(* IEC 61131-3 sources: TetherPLC/tests/compat (part 4) *)

(* ---- tc3_eventlog_case.st ---- *)
// tc3_eventlog_case.st — e2e for tc3_eventlog (tplc-eventlog).
PROGRAM tc3_eventlog_case
VAR
    msg : FB_TcMessage;
    alm : FB_TcAlarm;
    qry : FB_TcEventQuery;
    lg : FB_TcEventLogger;
    eb : FB_TcEventBase;
    ar : FB_TcArguments;
    si : FB_TcSourceInfo;
    st : INT;
    mask AT %QD0 : UDINT;
    diag AT %QD4 : UDINT;
END_VAR
    diag := st;
    IF st = 0 THEN
        mask := 0;
        msg.nEventClass := 7; msg.nEventId := 42;
        msg.sText := 'pump on'; msg.nCmd := 1;  // send INFO
        st := 1;
    ELSIF st = 1 THEN
        IF msg.bDone AND msg.hEvent <> 0 THEN mask := mask OR 1; END_IF;
        msg.nCmd := 0;
        alm.nEventClass := 7; alm.nEventId := 99;
        alm.nSeverity := 3; alm.sText := 'temp high';
        st := 2;
    ELSIF st = 2 THEN
        alm.nCmd := 1;                          // raise alarm
        st := 3;
    ELSIF st = 3 THEN
        IF alm.bDone AND alm.bActive AND alm.nState = 1 THEN
            mask := mask OR 2;
        END_IF;
        alm.nCmd := 0;
        st := 4;
    ELSIF st = 4 THEN
        alm.nCmd := 2;                          // clear
        st := 5;
    ELSIF st = 5 THEN
        IF alm.bDone AND alm.nState = 2 AND alm.bActive THEN
            mask := mask OR 4;
        END_IF;
        alm.nCmd := 0;
        st := 6;
    ELSIF st = 6 THEN
        qry.nId := alm.hEvent; qry.nCmd := 4;  // query the entry
        st := 7;
    ELSIF st = 7 THEN
        IF qry.bDone AND qry.nState = 2 AND qry.nSeverity = 3
           AND qry.nEventId = 99 THEN
            mask := mask OR 8;
        END_IF;
        qry.nCmd := 0;
        st := 8;
    ELSIF st = 8 THEN
        alm.nCmd := 3;                          // confirm
        st := 9;
    ELSIF st = 9 THEN
        IF alm.bDone AND NOT alm.bActive THEN mask := mask OR 16; END_IF;
        alm.nCmd := 0;
        st := 10;
    ELSIF st = 10 THEN
        // wrong-state op must error: query the released id
        qry.nId := 255; qry.nCmd := 4;
        st := 11;
    ELSIF st = 11 THEN
        IF qry.bError THEN mask := mask OR 32; END_IF;
        qry.nCmd := 0;
        st := 12;
    ELSIF st = 12 THEN
        qry.nCmd := 5;                          // stats
        st := 13;
    ELSIF st = 13 THEN
        IF qry.bDone AND qry.nRaised = 2 AND qry.nCleared = 1
           AND qry.nConfirmed = 1 AND qry.nLive = 1 THEN
            mask := mask OR 64;
        END_IF;
        qry.nCmd := 0;
        st := 14;
    ELSIF st = 14 THEN
        // second alarm for the aggregate/logger surface
        alm.nEventClass := 8; alm.nEventId := 77;
        alm.nSeverity := 3; alm.sText := 'overtemp';
        alm.nCmd := 1;
        lg.nFilterClass := 8; lg.nFilterEid := 0;
        st := 15;
    ELSIF st = 15 THEN
        IF alm.bDone THEN mask := mask OR 128; END_IF;
        alm.nCmd := 0;
        lg.nCmd := 7;                           // IsAlarmRaised
        st := 16;
    ELSIF st = 16 THEN
        lg.nCmd := 0;
        IF lg.bFound AND lg.nEidOut = 77 AND lg.nState = 1 THEN
            mask := mask OR 256;
        END_IF;
        st := 17;
    ELSIF st = 17 THEN
        lg.nCmd := 8;                           // GetAlarm
        st := 18;
    ELSIF st = 18 THEN
        lg.nCmd := 0;
        IF lg.bFound AND FIND(lg.sTextOut, 'overtemp') > 0 THEN
            mask := mask OR 512;
        END_IF;
        // EqualsToEventEntry against journal id 2
        eb.EventClass := 8; eb.EventId := 77;
        eb.Severity := 3; eb.Text := 'overtemp';
        eb.cEntryId := 2; eb.nCmd := 3;
        st := 19;
    ELSIF st = 19 THEN
        eb.nCmd := 0;
        IF eb.bEqual THEN mask := mask OR 1024; END_IF;
        lg.nCmd := 9;                           // ExportLoggedEvents
        st := 20;
    ELSIF st = 20 THEN
        lg.nCmd := 0;
        IF LEN(lg.sExport) > 0
           AND FIND(lg.sExport, ';') > 0
           AND FIND(lg.sExport, 'overtemp') > 0 THEN
            mask := mask OR 2048;
        END_IF;
        st := 21;
    ELSIF st = 21 THEN
        lg.nCmd := 2;                           // ClearAlarms (class 8)
        st := 22;
    ELSIF st = 22 THEN
        lg.nCmd := 0;
        IF lg.nCount = 1 THEN mask := mask OR 4096; END_IF;
        st := 23;
    ELSIF st = 23 THEN
        lg.nCmd := 5;                           // ConfirmAlarms
        st := 24;
    ELSIF st = 24 THEN
        lg.nCmd := 0;
        IF lg.nCount = 1 THEN mask := mask OR 8192; END_IF;
        // third alarm for the *All* variants
        alm.nEventClass := 8; alm.nEventId := 78;
        alm.nSeverity := 3; alm.sText := 'vibration';
        alm.nCmd := 1;
        st := 25;
    ELSIF st = 25 THEN
        IF alm.bDone THEN mask := mask OR 16384; END_IF;
        alm.nCmd := 0;
        lg.nCmd := 3;                           // ClearAllAlarms
        st := 26;
    ELSIF st = 26 THEN
        lg.nCmd := 0;
        IF lg.nCount >= 1 THEN mask := mask OR 32768; END_IF;
        st := 27;
    ELSIF st = 27 THEN
        lg.nCmd := 6;                           // ConfirmAllAlarms
        st := 28;
    ELSIF st = 28 THEN
        lg.nCmd := 0;
        IF lg.nCount >= 1 THEN mask := mask OR 65536; END_IF;
        st := 29;
    ELSIF st = 29 THEN
        lg.nCmd := 4;                           // ClearLoggedEvents
        st := 30;
    ELSIF st = 30 THEN
        lg.nCmd := 0;
        IF lg.nCount >= 1 THEN mask := mask OR 131072; END_IF;
        // FB_TcEventBase comparisons + text requests
        eb.EventClass := 8; eb.EventId := 77;
        eb.Severity := 3; eb.Text := 'overtemp';
        eb.cClass := 8; eb.cId := 77; eb.cSev := 3;
        eb.cText := 'overtemp'; eb.nCmd := 1;   // EqualsTo
        st := 31;
    ELSIF st = 31 THEN
        eb.nCmd := 0;
        IF eb.bEqual THEN mask := mask OR 262144; END_IF;
        st := 32;
    ELSIF st = 32 THEN
        eb.nCmd := 2;                           // EqualsToEventClass
        st := 33;
    ELSIF st = 33 THEN
        eb.nCmd := 0;
        IF eb.bEqual THEN mask := mask OR 524288; END_IF;
        st := 34;
    ELSIF st = 34 THEN
        eb.nCmd := 5;                           // RequestEventClassName
        st := 35;
    ELSIF st = 35 THEN
        eb.nCmd := 0;
        IF FIND(eb.sOut, '8') = 1 THEN mask := mask OR 1048576; END_IF;
        st := 36;
    ELSIF st = 36 THEN
        eb.nCmd := 6;                           // RequestEventText
        st := 37;
    ELSIF st = 37 THEN
        eb.nCmd := 0;
        IF FIND(eb.sOut, 'overtemp') = 1 THEN
            mask := mask OR 2097152;
        END_IF;
        ar.nInt := 5; ar.nCmd := 1;             // AddInt
        st := 38;
    ELSIF st = 38 THEN
        ar.nCmd := 0;
        st := 39;
    ELSIF st = 39 THEN
        IF ar.nCount = 1 THEN mask := mask OR 4194304; END_IF;
        ar.sArg := 'hi'; ar.nCmd := 3;          // AddString
        st := 40;
    ELSIF st = 40 THEN
        ar.nCmd := 0;
        st := 41;
    ELSIF st = 41 THEN
        IF ar.nCount = 2 THEN mask := mask OR 8388608; END_IF;
        si.Name := 'main'; si.nCmd := 1;        // ExtendName
        st := 42;
    ELSIF st = 42 THEN
        si.nCmd := 0;
        IF si.Extended THEN mask := mask OR 16777216; END_IF;
        st := 43;
    ELSIF st = 43 THEN
        ar.nCmd := 5;                           // Clear args
        st := 44;
    ELSIF st = 44 THEN
        ar.nCmd := 0;
        st := 45;
    ELSIF st = 45 THEN
        IF ar.bEmpty THEN mask := mask OR 33554432; END_IF;
        st := 46;
    END_IF;
    msg(); alm(); qry(); lg(); eb(); ar(); si();
END_PROGRAM

(* ---- tc3_ftp_case.st ---- *)
PROGRAM Tc3FtpCase
VAR
    mask      AT %QD0   : DINT;
    st        : INT;
    conn      : FB_FTP_Connect;
    connBad   : FB_FTP_Connect;
    sz        : FB_FTP_Cmd;
    mkd       : FB_FTP_MkDir;
    dl        : FB_FTP_Download;
    ls        : FB_FTP_List;
    up        : FB_FTP_Upload;
    szUp      : FB_FTP_Cmd;
    fex       : FB_FTP_FileExists;
    dex       : FB_FTP_DirExists;
    rn        : FB_FTP_Rename;
    acc       : ARRAY[0..1023] OF BYTE;
    accLen    : UDINT;
    i         : UDINT;
    upData    : ARRAY[0..511] OF BYTE;
END_VAR

// autonomous FTP sequence against tests/compat/ftp_test_peer.py
// (TCP 2121, PASV). The peer serves /data.txt (68B), /bin.dat,
// dirs / and /pub. Each state's bExecute is high only while st
// equals its index, giving every FB one rising edge; bDone
// advances the machine.
upData[0] := 16#50; upData[1] := 16#4C; upData[2] := 16#43;   // 'P','L','C'
upData[3] := 16#20; upData[4] := 16#75; upData[5] := 16#70;   // ' ','u','p'
// "PLC upload payload 12345" = 24 bytes
upData[6] := 16#6C; upData[7] := 16#6F; upData[8] := 16#61;
upData[9] := 16#64; upData[10] := 16#20; upData[11] := 16#70;
upData[12] := 16#61; upData[13] := 16#79; upData[14] := 16#6C;
upData[15] := 16#6F; upData[16] := 16#61; upData[17] := 16#64;
upData[18] := 16#20; upData[19] := 16#31; upData[20] := 16#32;
upData[21] := 16#33; upData[22] := 16#34; upData[23] := 16#35;

conn(sHost := '127.0.0.1', nPort := 2121, sUser := 'u', sPass := 'p',
     bExecute := st = 0, bClose := st = 11, tTimeout := T#5S);
connBad(sHost := '127.0.0.1', nPort := 21999, sUser := 'u', sPass := 'p',
        bExecute := st = 10, bClose := FALSE, tTimeout := T#3S);
sz(nConnHandle := conn.nConnHandle, sCmd := 'SIZE /data.txt',
   bExecute := st = 1, tTimeout := T#3S);
mkd(nConnHandle := conn.nConnHandle, sPath := '/newdir',
    bExecute := st = 2, tTimeout := T#3S);
dl(nConnHandle := conn.nConnHandle, sRemotePath := '/data.txt',
   bExecute := st = 3, tTimeout := T#10S);
ls(nConnHandle := conn.nConnHandle, sRemotePath := '/',
   bExecute := st = 4, tTimeout := T#10S);
up(nConnHandle := conn.nConnHandle, sRemotePath := '/up.bin',
   nLen := 24, DATA := upData, bExecute := st = 5, tTimeout := T#10S);
szUp(nConnHandle := conn.nConnHandle, sCmd := 'SIZE /up.bin',
     bExecute := st = 6, tTimeout := T#3S);
fex(nConnHandle := conn.nConnHandle, sPath := '/data.txt',
    bExecute := st = 7, tTimeout := T#3S);
dex(nConnHandle := conn.nConnHandle, sPath := '/pub',
    bExecute := st = 8, tTimeout := T#10S);
rn(nConnHandle := conn.nConnHandle, sOldPath := '/data.txt',
   sNewPath := '/renamed.txt', bExecute := st = 9, tTimeout := T#10S);

// accumulate download chunks every scan while st = 3
IF dl.nChunk > 0 AND accLen + dl.nChunk <= 1024 THEN
    FOR i := 0 TO dl.nChunk - 1 DO
        acc[accLen + i] := dl.DATA[i];
    END_FOR;
    accLen := accLen + dl.nChunk;
END_IF;

IF st = 0 AND conn.bDone THEN
    // connect -> login completes, handle issued
    IF conn.nStatus = 1 AND conn.nConnHandle <> 0 AND
       conn.nErrId = 0 THEN
        mask := mask + 1;
    END_IF;
    st := 1;
ELSIF st = 1 AND sz.bDone THEN
    // SIZE /data.txt -> 213, text "68"
    IF sz.nStatus = 1 AND sz.nRespCode = 213 AND
       sz.sText = '68' THEN
        mask := mask + 2;
    END_IF;
    st := 2;
ELSIF st = 2 AND mkd.bDone THEN
    // MKD /newdir -> 257
    IF mkd.nStatus = 1 AND mkd.nRespCode = 257 THEN
        mask := mask + 4;
    END_IF;
    st := 3;
ELSIF st = 3 AND dl.bDone THEN
    // RETR /data.txt -> 68 bytes "Hello FTP World!\n"x4
    IF dl.nStatus = 1 AND dl.nTotal = 68 AND accLen = 68 AND
       acc[0] = 16#48 AND acc[16] = 16#0A THEN
        mask := mask + 8;
    END_IF;
    st := 4;
ELSIF st = 4 AND ls.bDone THEN
    // LIST / -> non-empty listing
    IF ls.nStatus = 1 AND ls.nTotal > 0 THEN
        mask := mask + 16;
    END_IF;
    st := 5;
ELSIF st = 5 AND up.bDone THEN
    // STOR /up.bin -> 226
    IF up.nStatus = 1 AND up.nRespCode = 226 THEN
        mask := mask + 32;
    END_IF;
    st := 6;
ELSIF st = 6 AND szUp.bDone THEN
    // SIZE /up.bin -> 213 "24"
    IF szUp.nStatus = 1 AND szUp.nRespCode = 213 AND
       szUp.sText = '24' THEN
        mask := mask + 64;
    END_IF;
    st := 7;
ELSIF st = 7 AND fex.bDone THEN
    // FileExists /data.txt -> SIZE 213
    IF fex.bExists AND fex.nRespCode = 213 THEN
        mask := mask + 128;
    END_IF;
    st := 8;
ELSIF st = 8 AND dex.bDone THEN
    // DirExists /pub -> LIST ok
    IF dex.bExists AND dex.nStatus = 1 THEN
        mask := mask + 256;
    END_IF;
    st := 9;
ELSIF st = 9 AND rn.bDone THEN
    // Rename /data.txt -> /renamed.txt: RNFR 350 + RNTO 250
    IF rn.nStatus = 1 AND rn.nRespCode = 250 AND NOT rn.bError THEN
        mask := mask + 512;
    END_IF;
    st := 10;
ELSIF st = 10 AND connBad.bDone THEN
    // refused connect -> STATUS 2
    IF connBad.nStatus = 2 THEN
        mask := mask + 1024;
    END_IF;
    st := 11;
ELSIF st = 11 AND conn.bDone THEN
    // CLOSE -> session torn down
    IF conn.nConnHandle = 0 THEN
        mask := mask + 2048;
    END_IF;
    st := 12;
END_IF;
END_PROGRAM

(* ---- tc3_iec870_case.st ---- *)
PROGRAM Tc3Iec870Case
VAR
    mask      AT %QD0   : DINT;
    st        : INT;
    i2        : INT;
    conn      : FB_IEC870_5_104Master;
    connBad   : FB_IEC870_5_104Master;
    snd       : FB_IEC870_SendAsdu;
    snd2      : FB_IEC870_SendAsdu;
    snd3      : FB_IEC870_SendAsdu;
    rcv       : FB_IEC870_RecvAsdu;
    pay1      : ARRAY[0..239] OF BYTE;
    pay2      : ARRAY[0..239] OF BYTE;
    pay3      : ARRAY[0..239] OF BYTE;
    gotSp     : BOOL;
    gotMe     : BOOL;
    gotCs     : BOOL;
    gotSc     : BOOL;
    // helper-test vars
    o64       : ARRAY[0..6] OF BYTE;
    tenc      : SYSTEMTIME_TO_CP56Time2a;
    tdec      : CP56Time2a_TO_SYSTEMTIME;
    hY        : UDINT;
    hMo       : UDINT;
    hD        : UDINT;
    hH        : UDINT;
    hMi       : UDINT;
    hS        : UDINT;
    hMs       : UDINT;
    hbIV      : BOOL;
    hbSU      : BOOL;
    hVer      : UDINT;
    hCot      : STRING[31];
    hTid      : STRING[31];
    hIoa      : UDINT;
    hSpi      : BOOL;
    hDpi      : UDINT;
    hVti      : UDINT;
END_VAR

// autonomous IEC 60870-5-104 exchange against
// tests/compat/iec870_test_peer.py (TCP 2480). The peer is a
// slave: STARTDT handshake, then answers C_IC_NA_1 with
// M_SP_NA_1 + M_ME_NA_1, echoes C_CS_NA_1, answers C_SC_NA_1
// with an act-con. rcv() runs every scan (consume-on-read);
// each send gets one EXEC edge via its own st step.
rcv(nConnHandle := conn.nConnHandle);
IF rcv.bDone THEN
    // M_SP_NA_1: type1 vsq1 cot3 ca1 payload = IOA(3)+SPI(1)
    IF rcv.nTypeId = 1 AND rcv.nLen = 4 AND
       rcv.pPayload[2] = 1 AND rcv.pPayload[3] = 1 THEN
        gotSp := TRUE;
    END_IF;
    // M_ME_NA_1: type9 payload = IOA(3)+int16+QDS = 6 bytes
    IF rcv.nTypeId = 9 AND rcv.nLen = 6 AND
       rcv.pPayload[2] = 2 AND rcv.pPayload[3] = 16#34 AND
       rcv.pPayload[4] = 16#12 AND rcv.pPayload[5] = 0 THEN
        gotMe := TRUE;
    END_IF;
    IF rcv.nTypeId = 103 THEN
        gotCs := TRUE;
    END_IF;
    IF rcv.nTypeId = 45 THEN
        gotSc := TRUE;
    END_IF;
END_IF;

conn(sHost := '127.0.0.1', nPort := 2480, nCA_Size := 2,
     nCOT_Size := 2, bExecute := st = 0, bClose := st = 10,
     tTimeout := T#3S);
connBad(sHost := '127.0.0.1', nPort := 19999,
        bExecute := st = 8, bClose := FALSE, tTimeout := T#3S);

// payload staging
// pay1: interrogation C_IC_NA_1 has no info objects (len 0)
// pay2: C_CS_NA_1 clock sync, CP56Time2a = 13:45:30.250
// octets0-1 = sec*1000+ms = 30250 -> LE16 0x762A = 42,118
pay2[0] := 42; pay2[1] := 118;
pay2[2] := 45;                  // minute=45
pay2[3] := 13;                  // hour=13
pay2[4] := 15;                  // day=15
pay2[5] := 6;                   // month=6
pay2[6] := 124;                 // year-1900 = 2024-1900 = 124
// pay3: C_SC_NA_1 single command IOA=5, SCS=on -> 4 bytes
pay3[0] := 0; pay3[1] := 0; pay3[2] := 5; pay3[3] := 16#80;

snd(nConnHandle := conn.nConnHandle, nTypeId := 100, nVSQ := 0,
    nCOT := 5, nCA := 1, nLen := 0, pPayload := pay1,
    bExecute := st = 1);
snd2(nConnHandle := conn.nConnHandle, nTypeId := 103, nVSQ := 0,
     nCOT := 6, nCA := 1, nLen := 7, pPayload := pay2,
     bExecute := st = 4);
snd3(nConnHandle := conn.nConnHandle, nTypeId := 45, nVSQ := 1,
     nCOT := 6, nCA := 1, nLen := 4, pPayload := pay3,
     bExecute := st = 6);

IF st = 0 AND conn.bDone THEN
    IF conn.nStatus = 1 AND conn.nConnHandle <> 0 AND
       conn.nSubState = 3 AND conn.nErrId = 0 THEN
        mask := mask + 1;
    END_IF;
    st := 1;
ELSIF st = 1 AND snd.bDone THEN
    IF snd.nStatus = 1 AND snd.nErrId = 0 THEN
        mask := mask + 2;
    END_IF;
    st := 2;
ELSIF st = 2 AND gotSp AND gotMe THEN
    mask := mask + 4;
    st := 3;
ELSIF st = 3 THEN
    st := 4;
ELSIF st = 4 AND snd2.bDone THEN
    IF snd2.nStatus = 1 AND snd2.nErrId = 0 THEN
        mask := mask + 8;
    END_IF;
    st := 5;
ELSIF st = 5 AND gotCs THEN
    mask := mask + 16;
    st := 6;
ELSIF st = 6 AND snd3.bDone THEN
    IF snd3.nStatus = 1 AND snd3.nErrId = 0 THEN
        mask := mask + 32;
    END_IF;
    st := 7;
ELSIF st = 7 AND gotSc THEN
    mask := mask + 64;
    st := 8;
ELSIF st = 8 AND connBad.bDone THEN
    IF connBad.nStatus = 2 THEN
        mask := mask + 128;
    END_IF;
    st := 9;
ELSIF st = 9 THEN
    // pure-helper checks (single scan)
    // CP56Time2a roundtrip: encode 2024-06-15 13:45:30.250.
    // FB VAR_OUTPUT stays on the instance; copy pTime -> o64.
    tenc(nYear := 2024, nMonth := 6, nDay := 15,
         nHour := 13, nMinute := 45, nSecond := 30, nMs := 250,
         bIV := FALSE, bSU := FALSE);
    i2 := 0;
    WHILE i2 < 7 DO
        o64[i2] := tenc.pTime[i2];
        i2 := i2 + 1;
    END_WHILE;
    tdec(pTime := o64);
    hY := tdec.nYear; hMo := tdec.nMonth; hD := tdec.nDay;
    hH := tdec.nHour; hMi := tdec.nMinute; hS := tdec.nSecond;
    hMs := tdec.nMs; hbIV := tdec.bIV; hbSU := tdec.bSU;
    IF hY = 2024 AND hMo = 6 AND hD = 15 AND hH = 13 AND
       hMi = 45 AND hS = 30 AND hMs = 250 AND NOT hbIV THEN
        mask := mask + 256;
    END_IF;
    hCot := ASDU101COT_TO_STRING(3);
    hTid := ASDU101TYPEID_TO_STRING(9);
    IF hCot = 'SPONTANEOUS' AND hTid = 'M_ME_NA_1' THEN
        mask := mask + 512;
    END_IF;
    hIoa := CP24IOA_TO_DWORD(0, 0, 5);
    hSpi := F_iecGetSPI(1);
    hDpi := F_iecGetDPI(2);
    hVti := F_iecIncVTI(32767);
    hVer := GetIec870_Version();
    IF hIoa = 5 AND hSpi AND hDpi = 2 AND hVti = 0 AND
       hVer = 16#0100 THEN
        mask := mask + 1024;
    END_IF;
    st := 10;
ELSIF st = 10 THEN
    // bClose := st = 10 gave one rising edge -> session closed
    IF conn.nConnHandle = 0 THEN
        mask := mask + 2048;
        st := 11;
    END_IF;
END_IF;

END_PROGRAM

(* ---- tc3_jsonxml_case.st ---- *)
// tc3_jsonxml_case.st — e2e for tc3_jsonxml (pure-ST JSON).
// Builds a flat JSON object with FB_JsonSaxWriter, checks the
// text shape with FIND (string equality is not usable here),
// then parses it back with FB_JsonSaxReader.
PROGRAM tc3_jsonxml_case
VAR
    w : FB_JsonSaxWriter;
    r : FB_JsonSaxReader;
    doc : STRING[255];
    st : INT;
    mask AT %QD0 : UDINT;
    diag AT %QD4 : UDINT;
END_VAR
    diag := st;
    IF st = 0 THEN
        mask := 0;
        w.nCmd := 1;                        // Begin
        st := 1;
    ELSIF st = 1 THEN
        w.nCmd := 0;
        w.sKey := 'sp'; w.fReal := 12.5;
        st := 2;
    ELSIF st = 2 THEN
        w.nCmd := 4;                        // AddReal sp
        st := 3;
    ELSIF st = 3 THEN
        w.nCmd := 0;
        w.sKey := 'n'; w.nInt := 7;
        st := 4;
    ELSIF st = 4 THEN
        w.nCmd := 3;                        // AddInt n
        st := 5;
    ELSIF st = 5 THEN
        w.nCmd := 0;
        w.sKey := 'ok'; w.bBool := TRUE;
        st := 6;
    ELSIF st = 6 THEN
        w.nCmd := 5;                        // AddBool ok
        st := 7;
    ELSIF st = 7 THEN
        w.nCmd := 0;
        w.sKey := 's'; w.sVal := 'abc';
        st := 8;
    ELSIF st = 8 THEN
        w.nCmd := 2;                        // AddString s
        st := 9;
    ELSIF st = 9 THEN
        w.nCmd := 0;
        w.sKey := 'z';
        st := 10;
    ELSIF st = 10 THEN
        w.nCmd := 6;                        // AddNull z
        st := 11;
    ELSIF st = 11 THEN
        w.nCmd := 0;                        // clear so End sees an edge
        st := 12;
    ELSIF st = 12 THEN
        w.nCmd := 7;                        // End
        st := 13;
    ELSIF st = 13 THEN
        w.nCmd := 0;
        doc := w.sDoc;
        // shape checks (FIND, not equality)
        IF FIND(doc, '{"sp":12.500') = 1 THEN mask := mask OR 1; END_IF;
        IF FIND(doc, ',"n":7') > 0 THEN mask := mask OR 2; END_IF;
        IF FIND(doc, ',"ok":true') > 0 THEN mask := mask OR 4; END_IF;
        IF FIND(doc, ',"s":"abc"') > 0 THEN mask := mask OR 8; END_IF;
        IF FIND(doc, ',"z":null}') > 0 THEN mask := mask OR 16; END_IF;
        r.sIn := doc;
        st := 14;
    ELSIF st = 14 THEN
        r.nCmd := 1;                        // Load
        st := 15;
    ELSIF st = 15 THEN
        r.nCmd := 0;
        r.sKey := 'n';
        st := 16;
    ELSIF st = 16 THEN
        r.nCmd := 3;                        // GetInt n
        st := 17;
    ELSIF st = 17 THEN
        r.nCmd := 0;
        IF r.bDone AND r.nOut = 7 THEN mask := mask OR 32; END_IF;
        r.sKey := 'sp';
        st := 18;
    ELSIF st = 18 THEN
        r.nCmd := 4;                        // GetReal sp
        st := 19;
    ELSIF st = 19 THEN
        r.nCmd := 0;
        IF r.bDone AND r.fOut = 12.5 THEN mask := mask OR 64; END_IF;
        r.sKey := 'ok';
        st := 20;
    ELSIF st = 20 THEN
        r.nCmd := 5;                        // GetBool ok
        st := 21;
    ELSIF st = 21 THEN
        r.nCmd := 0;
        IF r.bDone AND r.bOut THEN mask := mask OR 128; END_IF;
        r.sKey := 's';
        st := 22;
    ELSIF st = 22 THEN
        r.nCmd := 2;                        // GetString s
        st := 23;
    ELSIF st = 23 THEN
        r.nCmd := 0;
        IF r.bDone AND FIND(r.sOut, 'abc') = 1 THEN mask := mask OR 256; END_IF;
        r.sKey := 'missing';
        st := 24;
    ELSIF st = 24 THEN
        r.nCmd := 2;                        // absent key -> error
        st := 25;
    ELSIF st = 25 THEN
        r.nCmd := 0;
        IF r.bError THEN mask := mask OR 512; END_IF;
        w.nCmd := 1;                        // Begin nested doc
        st := 27;
    ELSIF st = 27 THEN
        w.nCmd := 0;
        w.sKey := 'dev';
        st := 28;
    ELSIF st = 28 THEN
        w.nCmd := 9;                        // ObjBegin dev
        st := 29;
    ELSIF st = 29 THEN
        w.nCmd := 0;
        w.sKey := 'name'; w.sVal := 'ax1';
        st := 30;
    ELSIF st = 30 THEN
        w.nCmd := 2;                        // AddString name
        st := 31;
    ELSIF st = 31 THEN
        w.nCmd := 0;
        w.sKey := 'spd'; w.nInt := 2;
        st := 32;
    ELSIF st = 32 THEN
        w.nCmd := 3;                        // AddInt spd
        st := 33;
    ELSIF st = 33 THEN
        w.nCmd := 0;
        st := 34;
    ELSIF st = 34 THEN
        w.nCmd := 11;                       // EndAny -> close dev
        st := 35;
    ELSIF st = 35 THEN
        w.nCmd := 0;
        w.sKey := 'axes';
        st := 36;
    ELSIF st = 36 THEN
        w.nCmd := 10;                       // ArrBegin axes
        st := 37;
    ELSIF st = 37 THEN
        w.nCmd := 0;
        w.sKey := ''; w.nInt := 0;
        st := 38;
    ELSIF st = 38 THEN
        w.nCmd := 3;                        // array elem 0 (scalar)
        st := 39;
    ELSIF st = 39 THEN
        w.nCmd := 0;
        w.sKey := '';
        st := 40;
    ELSIF st = 40 THEN
        w.nCmd := 9;                        // ObjBegin elem object
        st := 41;
    ELSIF st = 41 THEN
        w.nCmd := 0;
        w.sKey := 'id'; w.nInt := 0;
        st := 42;
    ELSIF st = 42 THEN
        w.nCmd := 3;                        // AddInt id
        st := 43;
    ELSIF st = 43 THEN
        w.nCmd := 0;
        w.sKey := 'pos'; w.nInt := 100;
        st := 44;
    ELSIF st = 44 THEN
        w.nCmd := 3;                        // AddInt pos
        st := 45;
    ELSIF st = 45 THEN
        w.nCmd := 0;
        st := 46;
    ELSIF st = 46 THEN
        w.nCmd := 11;                       // EndAny -> close elem obj
        st := 47;
    ELSIF st = 47 THEN
        w.nCmd := 0;
        w.sKey := '';
        st := 48;
    ELSIF st = 48 THEN
        w.nCmd := 9;                        // ObjBegin elem 1
        st := 49;
    ELSIF st = 49 THEN
        w.nCmd := 0;
        w.sKey := 'id'; w.nInt := 1;
        st := 50;
    ELSIF st = 50 THEN
        w.nCmd := 3;
        st := 51;
    ELSIF st = 51 THEN
        w.nCmd := 0;
        w.sKey := 'pos'; w.nInt := 250;
        st := 52;
    ELSIF st = 52 THEN
        w.nCmd := 3;
        st := 53;
    ELSIF st = 53 THEN
        w.nCmd := 0;
        st := 54;
    ELSIF st = 54 THEN
        w.nCmd := 11;                       // EndAny -> close elem 1
        st := 55;
    ELSIF st = 55 THEN
        w.nCmd := 0;
        st := 56;
    ELSIF st = 56 THEN
        w.nCmd := 11;                       // EndAny -> close axes
        st := 57;
    ELSIF st = 57 THEN
        w.nCmd := 0;
        st := 58;
    ELSIF st = 58 THEN
        w.nCmd := 7;                        // End root
        st := 59;
    ELSIF st = 59 THEN
        w.nCmd := 0;
        doc := w.sDoc;
        IF FIND(doc, '"dev":{"name":"ax1","spd":2}') > 0
        THEN mask := mask OR 1024; END_IF;
        IF FIND(doc, ',"axes":[0,{"id":0,"pos":100}') > 0
        THEN mask := mask OR 2048; END_IF;
        IF FIND(doc, '{"id":1,"pos":250}]}') > 0
        THEN mask := mask OR 4096; END_IF;
        r.sIn := doc;
        st := 60;
    ELSIF st = 60 THEN
        r.nCmd := 1;                        // Load
        st := 61;
    ELSIF st = 61 THEN
        r.nCmd := 0;
        r.sKey := 'dev.spd';
        st := 62;
    ELSIF st = 62 THEN
        r.nCmd := 3;                        // GetInt dev.spd
        st := 63;
    ELSIF st = 63 THEN
        r.nCmd := 0;
        IF r.bDone AND r.nOut = 2 THEN mask := mask OR 8192; END_IF;
        r.sKey := 'axes.2.pos';
        st := 64;
    ELSIF st = 64 THEN
        r.nCmd := 3;                        // GetInt axes.2.pos
        st := 65;
    ELSIF st = 65 THEN
        r.nCmd := 0;
        IF r.bDone AND r.nOut = 250 THEN mask := mask OR 16384; END_IF;
        r.sKey := 'dev';
        st := 66;
    ELSIF st = 66 THEN
        r.nCmd := 2;                        // GetString dev -> raw obj
        st := 67;
    ELSIF st = 67 THEN
        r.nCmd := 0;
        IF r.bDone AND FIND(r.sOut, '"name"') > 0
        THEN mask := mask OR 32768; END_IF;
        r.sKey := 'axes.0.id';
        st := 68;
    ELSIF st = 68 THEN
        r.nCmd := 3;                        // GetInt axes.0.id -> elem1 obj? no:
        st := 69;                           // axes.0 is scalar 0, .id fails
    ELSIF st = 69 THEN
        r.nCmd := 0;
        // axes.0 is the scalar element 0; path 'axes.0.id' must fail
        IF r.bError THEN mask := mask OR 65536; END_IF;
        st := 70;
    END_IF;
    w(); r();
END_PROGRAM

(* ---- tc3_jsonxml_dom_case.st ---- *)
// tc3_jsonxml_dom_case.st — e2e for FB_JsonDomParser: load a
// document, query the tree, serialize, build a tree, error path.
// Every command needs a dedicated arm state + a reap state that
// clears nCmd (edge detect prev=0).
PROGRAM tc3_jsonxml_dom_case
VAR
    d : FB_JsonDomParser;
    doc : STRING[255];
    hR : UDINT;
    hDev : UDINT;
    hId : UDINT;
    hAx : UDINT;
    hA1 : UDINT;
    hF : UDINT;
    hN : UDINT;
    hR2 : UDINT;
    st : INT;
    mask AT %QD0 : UDINT;
    diag AT %QD4 : UDINT;
END_VAR
    diag := st;
    IF st = 0 THEN
        mask := 0;
        doc := CONCAT('{"name":"ax1","dev":{"id":7,"spd":1.5}',
            ',"axes":[1,2,3],"flag":true,"note":null}');
        d.sIn := doc;
        d.nCmd := 1;                        // Load
        st := 1;
    ELSIF st = 1 THEN                        // reap Load
        d.nCmd := 0;
        IF d.bDone THEN mask := mask OR 1; END_IF;
        st := 2;
    ELSIF st = 2 THEN                        // arm Root
        d.nCmd := 3;
        st := 3;
    ELSIF st = 3 THEN                        // reap Root
        d.nCmd := 0;
        hR := d.hOut;
        IF hR <> 0 THEN mask := mask OR 2; END_IF;
        st := 4;
    ELSIF st = 4 THEN                        // arm NodeType root
        d.hNode := hR;
        d.nCmd := 7;
        st := 5;
    ELSIF st = 5 THEN                        // reap
        d.nCmd := 0;
        IF d.nOut = 1 THEN mask := mask OR 4; END_IF;
        st := 6;
    ELSIF st = 6 THEN                        // arm ChildCount root
        d.hNode := hR;
        d.nCmd := 6;
        st := 7;
    ELSIF st = 7 THEN                        // reap
        d.nCmd := 0;
        IF d.nOut = 5 THEN mask := mask OR 8; END_IF;
        st := 8;
    ELSIF st = 8 THEN                        // arm ChildByName dev
        d.hNode := hR; d.sKey := 'dev';
        d.nCmd := 5;
        st := 9;
    ELSIF st = 9 THEN                        // reap -> hDev
        d.nCmd := 0;
        hDev := d.hOut;
        IF hDev <> 0 THEN mask := mask OR 16; END_IF;
        st := 10;
    ELSIF st = 10 THEN                       // arm NodeType dev
        d.hNode := hDev;
        d.nCmd := 7;
        st := 11;
    ELSIF st = 11 THEN                       // reap
        d.nCmd := 0;
        IF d.nOut = 1 THEN mask := mask OR 32; END_IF;
        st := 12;
    ELSIF st = 12 THEN                       // arm ChildByName id
        d.hNode := hDev; d.sKey := 'id';
        d.nCmd := 5;
        st := 13;
    ELSIF st = 13 THEN                       // reap -> hId
        d.nCmd := 0;
        hId := d.hOut;
        st := 14;
    ELSIF st = 14 THEN                       // arm NodeText id
        d.hNode := hId;
        d.nCmd := 9;
        st := 15;
    ELSIF st = 15 THEN                       // reap
        d.nCmd := 0;
        IF FIND(d.sOut, '7') = 1 THEN
            mask := mask OR 64;
        END_IF;
        st := 16;
    ELSIF st = 16 THEN                       // arm ChildByName axes
        d.hNode := hR; d.sKey := 'axes';
        d.nCmd := 5;
        st := 17;
    ELSIF st = 17 THEN                       // reap -> hAx
        d.nCmd := 0;
        hAx := d.hOut;
        st := 18;
    ELSIF st = 18 THEN                       // arm ChildCount axes
        d.hNode := hAx;
        d.nCmd := 6;
        st := 19;
    ELSIF st = 19 THEN                       // reap
        d.nCmd := 0;
        IF d.nOut = 3 THEN mask := mask OR 128; END_IF;
        st := 20;
    ELSIF st = 20 THEN                       // arm Child axes[1]
        d.hNode := hAx; d.nIdx := 1;
        d.nCmd := 4;
        st := 21;
    ELSIF st = 21 THEN                       // reap -> hA1
        d.nCmd := 0;
        hA1 := d.hOut;
        st := 22;
    ELSIF st = 22 THEN                       // arm NodeText axes[1]
        d.hNode := hA1;
        d.nCmd := 9;
        st := 23;
    ELSIF st = 23 THEN                       // reap
        d.nCmd := 0;
        IF FIND(d.sOut, '2') = 1 THEN
            mask := mask OR 256;
        END_IF;
        st := 24;
    ELSIF st = 24 THEN                       // arm ChildByName flag
        d.hNode := hR; d.sKey := 'flag';
        d.nCmd := 5;
        st := 25;
    ELSIF st = 25 THEN                       // reap -> hF
        d.nCmd := 0;
        hF := d.hOut;
        st := 26;
    ELSIF st = 26 THEN                       // arm NodeText flag
        d.hNode := hF;
        d.nCmd := 9;
        st := 27;
    ELSIF st = 27 THEN                       // reap
        d.nCmd := 0;
        IF FIND(d.sOut, 'true') = 1 THEN
            mask := mask OR 512;
        END_IF;
        st := 28;
    ELSIF st = 28 THEN                       // arm ChildByName note
        d.hNode := hR; d.sKey := 'note';
        d.nCmd := 5;
        st := 29;
    ELSIF st = 29 THEN                       // reap -> hN
        d.nCmd := 0;
        hN := d.hOut;
        st := 30;
    ELSIF st = 30 THEN                       // arm NodeType note
        d.hNode := hN;
        d.nCmd := 7;
        st := 31;
    ELSIF st = 31 THEN                       // reap
        d.nCmd := 0;
        IF d.nOut = 6 THEN mask := mask OR 1024; END_IF;
        st := 32;
    ELSIF st = 32 THEN                       // arm NodeKey dev
        d.hNode := hDev;
        d.nCmd := 8;
        st := 33;
    ELSIF st = 33 THEN                       // reap
        d.nCmd := 0;
        IF FIND(d.sOut, 'dev') = 1 THEN
            mask := mask OR 2048;
        END_IF;
        st := 34;
    ELSIF st = 34 THEN                       // arm ToJson whole doc
        d.hNode := 0;
        d.nCmd := 10;
        st := 35;
    ELSIF st = 35 THEN                       // reap
        d.nCmd := 0;
        IF FIND(d.sOut, '"name":"ax1"') > 0
           AND FIND(d.sOut, '"axes":[1,2,3]') > 0 THEN
            mask := mask OR 4096;
        END_IF;
        st := 36;
    ELSIF st = 36 THEN                       // arm Clear
        d.nCmd := 2;
        st := 37;
    ELSIF st = 37 THEN                       // reap Clear
        d.nCmd := 0;
        st := 38;
    ELSIF st = 38 THEN                       // arm AppendObject r
        d.hNode := 0; d.sKey := 'r';
        d.nCmd := 11;
        st := 39;
    ELSIF st = 39 THEN                       // reap -> hR2
        d.nCmd := 0;
        hR2 := d.hOut;
        st := 40;
    ELSIF st = 40 THEN                       // arm AppendString a=v
        d.hNode := hR2; d.sKey := 'a'; d.sVal := 'v';
        d.nCmd := 13;
        st := 41;
    ELSIF st = 41 THEN                       // reap
        d.nCmd := 0;
        st := 42;
    ELSIF st = 42 THEN                       // arm AppendInt n=42
        d.hNode := hR2; d.sKey := 'n'; d.nInt := 42;
        d.nCmd := 14;
        st := 43;
    ELSIF st = 43 THEN                       // reap
        d.nCmd := 0;
        st := 44;
    ELSIF st = 44 THEN                       // arm ToJson built tree
        d.hNode := 0;
        d.nCmd := 10;
        st := 45;
    ELSIF st = 45 THEN                       // reap
        d.nCmd := 0;
        IF FIND(d.sOut, '{"a":"v","n":42}') = 1 THEN
            mask := mask OR 8192;
        END_IF;
        st := 46;
    ELSIF st = 46 THEN                       // arm malformed Load
        d.sIn := '{"a":}';
        d.nCmd := 1;
        st := 47;
    ELSIF st = 47 THEN                       // reap error
        d.nCmd := 0;
        IF d.bError THEN mask := mask OR 16384; END_IF;
        st := 48;
    END_IF;
    d();
END_PROGRAM

(* ---- tc3_jsonxml_pretty_case.st ---- *)
// tc3_jsonxml_pretty_case.st — e2e for FB_JsonSaxPrettyWriter:
// indented JSON output.  Every command needs a dedicated arm
// state and a reap state that clears nCmd (edge detect prev=0).
PROGRAM tc3_jsonxml_pretty_case
VAR
    pw : FB_JsonSaxPrettyWriter;
    st : INT;
    mask AT %QD0 : UDINT;
    diag AT %QD4 : UDINT;
END_VAR
    diag := st;
    IF st = 0 THEN
        mask := 0;
        pw.nInt := 2;
        pw.nCmd := 12;                       // SetIndent 2
        st := 1;
    ELSIF st = 1 THEN                        // reap
        pw.nCmd := 0;
        st := 2;
    ELSIF st = 2 THEN                        // arm Begin
        pw.nCmd := 1;
        st := 3;
    ELSIF st = 3 THEN                        // reap
        pw.nCmd := 0;
        st := 4;
    ELSIF st = 4 THEN                        // arm AddString name
        pw.sKey := 'name'; pw.sVal := 'ax1';
        pw.nCmd := 2;
        st := 5;
    ELSIF st = 5 THEN                        // reap
        pw.nCmd := 0;
        st := 6;
    ELSIF st = 6 THEN                        // arm ObjBegin dev
        pw.sKey := 'dev';
        pw.nCmd := 9;
        st := 7;
    ELSIF st = 7 THEN                        // reap
        pw.nCmd := 0;
        st := 8;
    ELSIF st = 8 THEN                        // arm AddInt id
        pw.sKey := 'id'; pw.nInt := 7;
        pw.nCmd := 3;
        st := 9;
    ELSIF st = 9 THEN                        // reap
        pw.nCmd := 0;
        st := 10;
    ELSIF st = 10 THEN                       // arm AddReal spd
        pw.sKey := 'spd'; pw.fReal := 1.5;
        pw.nCmd := 4;
        st := 11;
    ELSIF st = 11 THEN                       // reap
        pw.nCmd := 0;
        st := 12;
    ELSIF st = 12 THEN                       // arm AddBool en
        pw.sKey := 'en'; pw.bBool := TRUE;
        pw.nCmd := 5;
        st := 13;
    ELSIF st = 13 THEN                       // reap
        pw.nCmd := 0;
        st := 14;
    ELSIF st = 14 THEN                       // arm EndAny dev
        pw.nCmd := 11;
        st := 15;
    ELSIF st = 15 THEN                       // reap
        pw.nCmd := 0;
        st := 16;
    ELSIF st = 16 THEN                       // arm ArrBegin axes
        pw.sKey := 'axes';
        pw.nCmd := 10;
        st := 17;
    ELSIF st = 17 THEN                       // reap
        pw.nCmd := 0;
        st := 18;
    ELSIF st = 18 THEN                       // arm AddInt 1
        pw.nInt := 1;
        pw.nCmd := 3;
        st := 19;
    ELSIF st = 19 THEN                       // reap
        pw.nCmd := 0;
        st := 20;
    ELSIF st = 20 THEN                       // arm AddInt 2
        pw.nInt := 2;
        pw.nCmd := 3;
        st := 21;
    ELSIF st = 21 THEN                       // reap
        pw.nCmd := 0;
        st := 22;
    ELSIF st = 22 THEN                       // arm EndAny axes
        pw.nCmd := 11;
        st := 23;
    ELSIF st = 23 THEN                       // reap
        pw.nCmd := 0;
        st := 24;
    ELSIF st = 24 THEN                       // arm End root
        pw.nCmd := 7;
        st := 25;
    ELSIF st = 25 THEN                       // reap + checks
        pw.nCmd := 0;
        IF pw.bDone THEN mask := mask OR 1; END_IF;
        IF FIND(pw.sDoc, '"dev": {') > 0 THEN
            mask := mask OR 2;
        END_IF;
        IF FIND(pw.sDoc, '
    "id": 7') > 0 THEN
            mask := mask OR 4;
        END_IF;
        IF FIND(pw.sDoc, '"axes": [') > 0 THEN
            mask := mask OR 8;
        END_IF;
        IF FIND(pw.sDoc, '1.500') > 0 THEN
            mask := mask OR 16;
        END_IF;
        IF FIND(pw.sDoc, '
}') > 0 AND NOT pw.bError THEN
            mask := mask OR 32;
        END_IF;
        st := 26;
    END_IF;
    pw();
END_PROGRAM

(* ---- tc3_jsonxml_xml_case.st ---- *)
// tc3_jsonxml_xml_case.st — e2e for the XML half of tc3_jsonxml:
// FB_XmlDomParser load/query/serialize + build commands.
// Command FBs need a full scan with nCmd=0 between commands (edge
// detect on prev=0): every command gets a dedicated arm state, then
// a reap state that clears nCmd and reads the outputs.
PROGRAM tc3_jsonxml_xml_case
VAR
    x : FB_XmlDomParser;
    xdoc : STRING[1023];
    hRoot : UDINT;
    hDev : UDINT;
    hNm : UDINT;
    hPos : UDINT;
    hAx : UDINT;
    hTmp : UDINT;
    st : INT;
    mask AT %QD0 : UDINT;
    diag AT %QD4 : UDINT;
END_VAR
    diag := st;
    IF st = 0 THEN
        mask := 0;
        xdoc := CONCAT('<?xml version="1.0"?>',
            CONCAT('<root><dev id="ax1" unit="mm">',
            CONCAT('<name>motor</name><pos>100</pos></dev>',
            CONCAT('<axes><axis pos="1"/><axis pos="2"/>',
                   '<axis pos="3"/></axes></root>'))));
        x.sIn := xdoc; x.nCmd := 1;           // Load
        st := 1;
    // reap Load
    ELSIF st = 1 THEN
        x.nCmd := 0;
        IF x.bDone THEN mask := mask OR 1; END_IF;
        st := 2;
    // arm Root
    ELSIF st = 2 THEN
        x.nCmd := 3;
        st := 3;
    // reap Root
    ELSIF st = 3 THEN
        x.nCmd := 0;
        hRoot := x.hOut;
        IF hRoot <> 0 THEN mask := mask OR 2; END_IF;
        st := 4;
    // arm NodeName root
    ELSIF st = 4 THEN
        x.hNode := hRoot;
        x.nCmd := 6;
        st := 5;
    // reap NodeName
    ELSIF st = 5 THEN
        x.nCmd := 0;
        IF FIND(x.sOut, 'root') = 1 THEN
            mask := mask OR 4;
        END_IF;
        st := 6;
    // arm ChildByName dev
    ELSIF st = 6 THEN
        x.hNode := hRoot; x.sName := 'dev';
        x.nCmd := 5;
        st := 7;
    // reap -> hDev
    ELSIF st = 7 THEN
        x.nCmd := 0;
        hDev := x.hOut;
        IF hDev <> 0 THEN mask := mask OR 8; END_IF;
        st := 8;
    // arm AttrByName id
    ELSIF st = 8 THEN
        x.hNode := hDev; x.sName := 'id';
        x.nCmd := 10;
        st := 9;
    // reap attr id
    ELSIF st = 9 THEN
        x.nCmd := 0;
        IF FIND(x.sOut, 'ax1') = 1 THEN
            mask := mask OR 16;
        END_IF;
        st := 10;
    // arm AttrCount dev
    ELSIF st = 10 THEN
        x.hNode := hDev;
        x.nCmd := 8;
        st := 11;
    // reap AttrCount
    ELSIF st = 11 THEN
        x.nCmd := 0;
        IF x.nOut = 2 THEN mask := mask OR 32; END_IF;
        st := 12;
    // arm ChildByName name
    ELSIF st = 12 THEN
        x.hNode := hDev; x.sName := 'name';
        x.nCmd := 5;
        st := 13;
    // reap -> hNm
    ELSIF st = 13 THEN
        x.nCmd := 0;
        hNm := x.hOut;
        st := 14;
    // arm NodeText name
    ELSIF st = 14 THEN
        x.hNode := hNm;
        x.nCmd := 7;
        st := 15;
    // reap NodeText
    ELSIF st = 15 THEN
        x.nCmd := 0;
        IF FIND(x.sOut, 'motor') = 1 THEN
            mask := mask OR 64;
        END_IF;
        st := 16;
    // arm ChildByName pos
    ELSIF st = 16 THEN
        x.hNode := hDev; x.sName := 'pos';
        x.nCmd := 5;
        st := 17;
    // reap -> hPos
    ELSIF st = 17 THEN
        x.nCmd := 0;
        hPos := x.hOut;
        st := 18;
    // arm NodeText pos
    ELSIF st = 18 THEN
        x.hNode := hPos;
        x.nCmd := 7;
        st := 19;
    // reap NodeText pos
    ELSIF st = 19 THEN
        x.nCmd := 0;
        IF FIND(x.sOut, '100') = 1 THEN
            mask := mask OR 128;
        END_IF;
        st := 20;
    // arm ChildByName axes
    ELSIF st = 20 THEN
        x.hNode := hRoot; x.sName := 'axes';
        x.nCmd := 5;
        st := 21;
    // reap -> hAx
    ELSIF st = 21 THEN
        x.nCmd := 0;
        hAx := x.hOut;
        st := 22;
    // arm ChildCount axes
    ELSIF st = 22 THEN
        x.hNode := hAx;
        x.nCmd := 9;
        st := 23;
    // reap ChildCount
    ELSIF st = 23 THEN
        x.nCmd := 0;
        IF x.nOut = 3 THEN mask := mask OR 256; END_IF;
        st := 24;
    // arm Child axes[1] (0-based -> second axis)
    ELSIF st = 24 THEN
        x.hNode := hAx; x.nIdx := 1;
        x.nCmd := 4;
        st := 25;
    // reap -> hTmp
    ELSIF st = 25 THEN
        x.nCmd := 0;
        hTmp := x.hOut;
        st := 26;
    // arm AttrByName pos on axis2
    ELSIF st = 26 THEN
        x.hNode := hTmp; x.sName := 'pos';
        x.nCmd := 10;
        st := 27;
    // reap attr pos
    ELSIF st = 27 THEN
        x.nCmd := 0;
        IF FIND(x.sOut, '2') = 1 THEN
            mask := mask OR 512;
        END_IF;
        st := 28;
    // arm NodeXml dev
    ELSIF st = 28 THEN
        x.hNode := hDev;
        x.nCmd := 11;
        st := 29;
    // reap NodeXml
    ELSIF st = 29 THEN
        x.nCmd := 0;
        IF FIND(x.sOut, 'id="ax1"') > 0
           AND FIND(x.sOut, '<name>') > 0 THEN
            mask := mask OR 1024;
        END_IF;
        st := 30;
    // arm ToXml
    ELSIF st = 30 THEN
        x.hNode := 0;
        x.nCmd := 12;
        st := 31;
    // reap ToXml
    ELSIF st = 31 THEN
        x.nCmd := 0;
        IF FIND(x.sOut, '</root>') > 0
           AND FIND(x.sOut, '<axis') > 0 THEN
            mask := mask OR 2048;
        END_IF;
        st := 32;
    // arm Clear
    ELSIF st = 32 THEN
        x.nCmd := 2;
        st := 33;
    // reap Clear
    ELSIF st = 33 THEN
        x.nCmd := 0;
        st := 34;
    // arm AppendChild r under #doc
    ELSIF st = 34 THEN
        x.hNode := 0; x.sName := 'r';
        x.nCmd := 13;
        st := 35;
    // reap -> hRoot (new tree)
    ELSIF st = 35 THEN
        x.nCmd := 0;
        hRoot := x.hOut;
        st := 36;
    // arm AppendAttribute a=v on r
    ELSIF st = 36 THEN
        x.hNode := hRoot; x.sName := 'a'; x.sVal := 'v';
        x.nCmd := 14;
        st := 37;
    // reap attr
    ELSIF st = 37 THEN
        x.nCmd := 0;
        st := 38;
    // arm AppendChild c under r
    ELSIF st = 38 THEN
        x.hNode := hRoot; x.sName := 'c';
        x.nCmd := 13;
        st := 39;
    // reap -> hNm
    ELSIF st = 39 THEN
        x.nCmd := 0;
        hNm := x.hOut;
        st := 40;
    // arm AppendText hi on c
    ELSIF st = 40 THEN
        x.hNode := hNm; x.sVal := 'hi';
        x.nCmd := 15;
        st := 41;
    // reap text
    ELSIF st = 41 THEN
        x.nCmd := 0;
        st := 42;
    // arm ToXml of built tree
    ELSIF st = 42 THEN
        x.hNode := 0;
        x.nCmd := 12;
        st := 43;
    // reap ToXml
    ELSIF st = 43 THEN
        x.nCmd := 0;
        IF FIND(x.sOut, '<r a="v"><c>hi</c></r>') = 1 THEN
            mask := mask OR 4096;
        END_IF;
        st := 44;
    // arm malformed Load
    ELSIF st = 44 THEN
        x.sIn := '<a x></a>';
        x.nCmd := 1;
        st := 45;
    // reap error
    ELSIF st = 45 THEN
        x.nCmd := 0;
        IF x.bError THEN mask := mask OR 8192; END_IF;
        st := 46;
    END_IF;
    x();
END_PROGRAM

(* ---- tc3_mc2_ah_case.st ---- *)
// e2e for compat/tc3/tc3_mc2_ah.st — Tc3_MC2_AdvancedHoming:
// step search FBs (ref pulse, absolute switch, limit switch,
// block, block-lag), detection variants, finalizing FBs and a
// flying (passive) reference over a simulated axis.
// Mask bits (expected 0xFFFF):
//  0 axis created   1 powered        2 pos preset     3 refPulse
//  4 absSwitchDet   5 absSwitch      6 limitSwitch    7 block
//  8 blockDet       9 blockLag      10 homeDirect    11 finishHome
// 12 abortHome     13 flyingSwitch  14 errBadVel    15 errBadDir
PROGRAM Tc3Mc2AhCase
VAR
    mask   AT %QD0 : DINT;
    st     : INT;
    prevSt : INT;
    started: BOOL;
    pulse  : BOOL;

    ax     : FB_MotionAxis;
    rd     : FB_MotionAxis;
    axM    : UDINT;

    pwr    : MC_Power;
    sp     : MC_SetPosition;
    stp    : MC_Stop;
    mv     : MC_MoveVelocity;

    // homing FBs under test
    refPls : MC_StepReferencePulse;
    refPls2: MC_StepReferencePulse;
    refPls3: MC_StepReferencePulse;
    absDet : MC_StepAbsoluteSwitchDetection;
    absSw  : MC_StepAbsoluteSwitch;
    limSw  : MC_StepLimitSwitch;
    blk    : MC_StepBlock;
    blkDet : MC_StepBlockDetection;
    blkLag : MC_StepBlockLagBased;
    finH   : MC_FinishHoming;
    homeDir: MC_HomeDirect;
    abortH : MC_AbortHoming;
    flySw  : MC_StepReferenceFlyingSwitch;

    // shared MC_HomingParameter (flattened) state
    pStored : BOOL;
    pNcSMin : BOOL;  pNcSMax : BOOL;
    pNcSPosDiff : BOOL;  pNcSVeloDiff : BOOL;
    pNcAMin : BOOL;  pNcAMax : BOOL;
    pNcAPosDiff : BOOL;  pNcAVeloDiff : BOOL;
    pDrvSBip : LREAL;  pDrvSPos : LREAL;  pDrvSNeg : LREAL;
    pDrvABip : LREAL;  pDrvAPos : LREAL;  pDrvANeg : LREAL;

    // simulated reference signals (position-derived levels)
    dRef   : BOOL; dAbsD : BOOL; dAbsS : BOOL; dLim  : BOOL;
    dBlk   : BOOL; dBlkD : BOOL; dBlkL : BOOL; dHomeD : BOOL;
    dFin   : BOOL; dAbort: BOOL; dFly  : BOOL;
    sigZ   : BOOL;
    sigAbs : BOOL;
    sigLim : BOOL;
    sigFly : BOOL;

    posL   : LREAL;
    enSig  : BOOL;
    mvEx   : BOOL;
    spEx   : BOOL;
    stpEx  : BOOL;
    finEx  : BOOL;
    dirEx  : BOOL;
    abortEx: BOOL;
    flyEx  : BOOL;
    errEx  : BOOL;
    errEx2 : BOOL;
    refEx  : BOOL;
    absDetEx : BOOL;
    absSwEx  : BOOL;
    limSwEx  : BOOL;
    blkEx    : BOOL;
    blkDetEx : BOOL;
    blkLagEx : BOOL;
    homeDirEx: BOOL;
    errId1 : UDINT;
    errId2 : UDINT;
END_VAR

// ---- per-scan FB calls ----------------------------------------------
IF NOT started THEN
    pulse := TRUE; started := TRUE;
ELSIF st <> prevSt THEN
    pulse := TRUE;
ELSE
    pulse := FALSE;
END_IF;
prevSt := st;

IF axM <> 0 THEN
    rd.AXIS := axM; rd.OP := 6; rd();
END_IF;
posL := DINT_TO_LREAL(rd.POS_ACTUAL);

// reference signals derived from axis position
sigZ   := posL >= 5000.0;
sigAbs := posL >= 8000.0;
sigLim := posL <= -5000.0;
sigFly := posL >= 3000.0;

// execute pulses: launch stages, waits follow on the next stage
enSig := (st >= 1);
mvEx  := pulse AND (st = 38);
spEx  := pulse AND ((st = 2) OR (st = 6) OR (st = 10) OR (st = 14)
                    OR (st = 18) OR (st = 22) OR (st = 26));
stpEx := pulse AND (st = 42);
finEx := pulse AND (st = 33);
dirEx := pulse AND (st = 31);
abortEx := pulse AND (st = 35);
flyEx := pulse AND (st = 39);
errEx := pulse AND (st = 44);
errEx2 := pulse AND (st = 46);
refEx := pulse AND (st = 4);
absDetEx := pulse AND (st = 8);
absSwEx  := pulse AND (st = 12);
limSwEx  := pulse AND (st = 16);
blkEx    := pulse AND (st = 20);
blkDetEx := pulse AND (st = 24);
blkLagEx := pulse AND (st = 28);
homeDirEx:= dirEx;

pwr(Enable := enSig, Enable_Positive := TRUE, Enable_Negative := TRUE,
    Axis := axM);
sp(Execute := spEx, Position := 0, Mode := FALSE, Axis := axM);
stp(Execute := stpEx, Deceleration := 50000, Axis := axM);
mv(Execute := mvEx, ContinuousUpdate := FALSE, Velocity := 5000,
   Acceleration := 50000, Deceleration := 50000, Axis := axM);

// ---- homing FB calls (every scan; Execute is edge-driven inside) --
refPls(
       Execute := refEx,  Direction := 1,  SwitchMode := 3,
       RefLevel := sigZ,  Velocity := 20000.0,
       Acceleration := 50000.0,  Deceleration := 50000.0,  Jerk := 0.0,
       SetPosition := 100.0,  TimeLimit := T#0s,
       DistanceLimit := 50000.0,  TorqueLimit := 0.0,  BufferMode := 0,
       OptDisableDriveAccess := FALSE,
       OptEnableLagErrorDetection := FALSE,  Axis := axM,
       P_Stored := pStored,  P_NcSMin := pNcSMin,  P_NcSMax := pNcSMax,
       P_NcSPosDiff := pNcSPosDiff,  P_NcSVeloDiff := pNcSVeloDiff,
       P_NcAMin := pNcAMin,  P_NcAMax := pNcAMax,
       P_NcAPosDiff := pNcAPosDiff,  P_NcAVeloDiff := pNcAVeloDiff,
       P_DrvSBip := pDrvSBip,  P_DrvSPos := pDrvSPos,
       P_DrvSNeg := pDrvSNeg,  P_DrvABip := pDrvABip,
       P_DrvAPos := pDrvAPos,  P_DrvANeg := pDrvANeg);
absDet(
       Execute := absDetEx,  Direction := 3,  SwitchMode := 3,
       RefLevel := (posL <= -3000.0),  Velocity := 20000.0,
       Acceleration := 50000.0,  Deceleration := 50000.0,  Jerk := 0.0,
       TimeLimit := T#0s,  DistanceLimit := 50000.0,
       TorqueLimit := 0.0,  PositiveLimitSwitch := FALSE,
       NegativeLimitSwitch := FALSE,  BufferMode := 0,
       OptDisableDriveAccess := FALSE,
       OptEnableLagErrorDetection := FALSE,  Axis := axM,
       P_Stored := pStored,  P_NcSMin := pNcSMin,  P_NcSMax := pNcSMax,
       P_NcSPosDiff := pNcSPosDiff,  P_NcSVeloDiff := pNcSVeloDiff,
       P_NcAMin := pNcAMin,  P_NcAMax := pNcAMax,
       P_NcAPosDiff := pNcAPosDiff,  P_NcAVeloDiff := pNcAVeloDiff,
       P_DrvSBip := pDrvSBip,  P_DrvSPos := pDrvSPos,
       P_DrvSNeg := pDrvSNeg,  P_DrvABip := pDrvABip,
       P_DrvAPos := pDrvAPos,  P_DrvANeg := pDrvANeg);
absSw(
       Execute := absSwEx,  Direction := 1,  SwitchMode := 3,
       RefLevel := sigAbs,  Velocity := 20000.0,
       Acceleration := 50000.0,  Deceleration := 50000.0,  Jerk := 0.0,
       SetPosition := 500.0,  TimeLimit := T#0s,
       DistanceLimit := 50000.0,  TorqueLimit := 0.0,
       PositiveLimitSwitch := FALSE,  NegativeLimitSwitch := FALSE,
       BufferMode := 0,  OptDisableDriveAccess := FALSE,
       OptEnableLagErrorDetection := FALSE,  Axis := axM,
       P_Stored := pStored,  P_NcSMin := pNcSMin,  P_NcSMax := pNcSMax,
       P_NcSPosDiff := pNcSPosDiff,  P_NcSVeloDiff := pNcSVeloDiff,
       P_NcAMin := pNcAMin,  P_NcAMax := pNcAMax,
       P_NcAPosDiff := pNcAPosDiff,  P_NcAVeloDiff := pNcAVeloDiff,
       P_DrvSBip := pDrvSBip,  P_DrvSPos := pDrvSPos,
       P_DrvSNeg := pDrvSNeg,  P_DrvABip := pDrvABip,
       P_DrvAPos := pDrvAPos,  P_DrvANeg := pDrvANeg);
limSw(
       Execute := limSwEx,  Direction := 3,  LimitSwitchMode := 3,
       LimitSwitchLevel := sigLim,  Velocity := 20000.0,
       Acceleration := 50000.0,  Deceleration := 50000.0,  Jerk := 0.0,
       SetPosition := -500.0,  TimeLimit := T#0s,
       DistanceLimit := 50000.0,  TorqueLimit := 0.0,  BufferMode := 0,
       OptDisableDriveAccess := FALSE,
       OptEnableLagErrorDetection := FALSE,  Axis := axM,
       P_Stored := pStored,  P_NcSMin := pNcSMin,  P_NcSMax := pNcSMax,
       P_NcSPosDiff := pNcSPosDiff,  P_NcSVeloDiff := pNcSVeloDiff,
       P_NcAMin := pNcAMin,  P_NcAMax := pNcAMax,
       P_NcAPosDiff := pNcAPosDiff,  P_NcAVeloDiff := pNcAVeloDiff,
       P_DrvSBip := pDrvSBip,  P_DrvSPos := pDrvSPos,
       P_DrvSNeg := pDrvSNeg,  P_DrvABip := pDrvABip,
       P_DrvAPos := pDrvAPos,  P_DrvANeg := pDrvANeg);
blk(
       Execute := blkEx,  Direction := 1,  Velocity := 80000.0,
       Acceleration := 50000.0,  Deceleration := 50000.0,  Jerk := 0.0,
       SetPosition := 25000.0,  DetectionVelocityLimit := 800.0,
       DetectionVelocityTime := T#100ms,  TimeLimit := T#0s,
       DistanceLimit := 40000.0,  TorqueLimit := 0.0,
       TorqueTolerance := 0.0,  BufferMode := 0,
       OptDisableDriveAccess := FALSE,
       OptInstantLagReduction := FALSE,  Axis := axM,
       P_Stored := pStored,  P_NcSMin := pNcSMin,  P_NcSMax := pNcSMax,
       P_NcSPosDiff := pNcSPosDiff,  P_NcSVeloDiff := pNcSVeloDiff,
       P_NcAMin := pNcAMin,  P_NcAMax := pNcAMax,
       P_NcAPosDiff := pNcAPosDiff,  P_NcAVeloDiff := pNcAVeloDiff,
       P_DrvSBip := pDrvSBip,  P_DrvSPos := pDrvSPos,
       P_DrvSNeg := pDrvSNeg,  P_DrvABip := pDrvABip,
       P_DrvAPos := pDrvAPos,  P_DrvANeg := pDrvANeg);
blkDet(
       Execute := blkDetEx,  Direction := 3,  Velocity := 80000.0,
       Acceleration := 50000.0,  Deceleration := 50000.0,  Jerk := 0.0,
       DetectionVelocityLimit := 800.0,
       DetectionVelocityTime := T#100ms,  TimeLimit := T#0s,
       DistanceLimit := 40000.0,  TorqueLimit := 0.0,
       TorqueTolerance := 0.0,  BufferMode := 0,
       OptDisableDriveAccess := FALSE,
       OptInstantLagReduction := FALSE,  Axis := axM,
       P_Stored := pStored,  P_NcSMin := pNcSMin,  P_NcSMax := pNcSMax,
       P_NcSPosDiff := pNcSPosDiff,  P_NcSVeloDiff := pNcSVeloDiff,
       P_NcAMin := pNcAMin,  P_NcAMax := pNcAMax,
       P_NcAPosDiff := pNcAPosDiff,  P_NcAVeloDiff := pNcAVeloDiff,
       P_DrvSBip := pDrvSBip,  P_DrvSPos := pDrvSPos,
       P_DrvSNeg := pDrvSNeg,  P_DrvABip := pDrvABip,
       P_DrvAPos := pDrvAPos,  P_DrvANeg := pDrvANeg);
blkLag(
       Execute := blkLagEx,  Direction := 1,  Velocity := 80000.0,
       Acceleration := 50000.0,  Deceleration := 50000.0,  Jerk := 0.0,
       SetPosition := 20000.0,  DetectionVelocityLimit := 800.0,
       DetectionVelocityTime := T#100ms,  TimeLimit := T#0s,
       DistanceLimit := 40000.0,  TorqueLimit := 0.0,
       LagLimit := 1000.0,  BufferMode := 0,
       OptDisableDriveAccess := FALSE,
       OptInstantLagReduction := FALSE,  Axis := axM,
       P_Stored := pStored,  P_NcSMin := pNcSMin,  P_NcSMax := pNcSMax,
       P_NcSPosDiff := pNcSPosDiff,  P_NcSVeloDiff := pNcSVeloDiff,
       P_NcAMin := pNcAMin,  P_NcAMax := pNcAMax,
       P_NcAPosDiff := pNcAPosDiff,  P_NcAVeloDiff := pNcAVeloDiff,
       P_DrvSBip := pDrvSBip,  P_DrvSPos := pDrvSPos,
       P_DrvSNeg := pDrvSNeg,  P_DrvABip := pDrvABip,
       P_DrvAPos := pDrvAPos,  P_DrvANeg := pDrvANeg);
homeDir(
       Execute := homeDirEx,  SetPosition := 777.0,  BufferMode := 0,
       OptDisableDriveAccess := FALSE,  Axis := axM,
       P_Stored := pStored,  P_NcSMin := pNcSMin,  P_NcSMax := pNcSMax,
       P_NcSPosDiff := pNcSPosDiff,  P_NcSVeloDiff := pNcSVeloDiff,
       P_NcAMin := pNcAMin,  P_NcAMax := pNcAMax,
       P_NcAPosDiff := pNcAPosDiff,  P_NcAVeloDiff := pNcAVeloDiff,
       P_DrvSBip := pDrvSBip,  P_DrvSPos := pDrvSPos,
       P_DrvSNeg := pDrvSNeg,  P_DrvABip := pDrvABip,
       P_DrvAPos := pDrvAPos,  P_DrvANeg := pDrvANeg);
finH(
       Execute := finEx,  Distance := 500.0,  Velocity := 1000.0,
       Acceleration := 50000.0,  Deceleration := 50000.0,  Jerk := 0.0,
       BufferMode := 0,  OptDisableDriveAccess := FALSE,  Axis := axM,
       P_Stored := pStored,  P_NcSMin := pNcSMin,  P_NcSMax := pNcSMax,
       P_NcSPosDiff := pNcSPosDiff,  P_NcSVeloDiff := pNcSVeloDiff,
       P_NcAMin := pNcAMin,  P_NcAMax := pNcAMax,
       P_NcAPosDiff := pNcAPosDiff,  P_NcAVeloDiff := pNcAVeloDiff,
       P_DrvSBip := pDrvSBip,  P_DrvSPos := pDrvSPos,
       P_DrvSNeg := pDrvSNeg,  P_DrvABip := pDrvABip,
       P_DrvAPos := pDrvAPos,  P_DrvANeg := pDrvANeg);
abortH(
       Execute := abortEx,  OptDisableDriveAccess := FALSE,
       Axis := axM,  P_Stored := pStored,  P_NcSMin := pNcSMin,
       P_NcSMax := pNcSMax,  P_NcSPosDiff := pNcSPosDiff,
       P_NcSVeloDiff := pNcSVeloDiff,  P_NcAMin := pNcAMin,
       P_NcAMax := pNcAMax,  P_NcAPosDiff := pNcAPosDiff,
       P_NcAVeloDiff := pNcAVeloDiff,  P_DrvSBip := pDrvSBip,
       P_DrvSPos := pDrvSPos,  P_DrvSNeg := pDrvSNeg,
       P_DrvABip := pDrvABip,  P_DrvAPos := pDrvAPos,
       P_DrvANeg := pDrvANeg);
flySw(
       Execute := flyEx,  SwitchMode := 3,  RefLevel := sigFly,
       SetPosition := 4242.0,  TimeLimit := T#0s,
       DistanceLimit := 50000.0,  BufferMode := 0,  Axis := axM);
refPls2(
       Execute := errEx,  Direction := 1,  SwitchMode := 3,
       RefLevel := FALSE,  Velocity := 0.0,  Acceleration := 50000.0,
       Deceleration := 50000.0,  Jerk := 0.0,  SetPosition := 0.0,
       TimeLimit := T#0s,  DistanceLimit := 50000.0,
       TorqueLimit := 0.0,  BufferMode := 0,
       OptDisableDriveAccess := FALSE,
       OptEnableLagErrorDetection := FALSE,  Axis := axM,
       P_Stored := pStored,  P_NcSMin := pNcSMin,  P_NcSMax := pNcSMax,
       P_NcSPosDiff := pNcSPosDiff,  P_NcSVeloDiff := pNcSVeloDiff,
       P_NcAMin := pNcAMin,  P_NcAMax := pNcAMax,
       P_NcAPosDiff := pNcAPosDiff,  P_NcAVeloDiff := pNcAVeloDiff,
       P_DrvSBip := pDrvSBip,  P_DrvSPos := pDrvSPos,
       P_DrvSNeg := pDrvSNeg,  P_DrvABip := pDrvABip,
       P_DrvAPos := pDrvAPos,  P_DrvANeg := pDrvANeg);
refPls3(
       Execute := errEx2,  Direction := 9,  SwitchMode := 3,
       RefLevel := FALSE,  Velocity := 100.0,  Acceleration := 50000.0,
       Deceleration := 50000.0,  Jerk := 0.0,  SetPosition := 0.0,
       TimeLimit := T#0s,  DistanceLimit := 50000.0,
       TorqueLimit := 0.0,  BufferMode := 0,
       OptDisableDriveAccess := FALSE,
       OptEnableLagErrorDetection := FALSE,  Axis := axM,
       P_Stored := pStored,  P_NcSMin := pNcSMin,  P_NcSMax := pNcSMax,
       P_NcSPosDiff := pNcSPosDiff,  P_NcSVeloDiff := pNcSVeloDiff,
       P_NcAMin := pNcAMin,  P_NcAMax := pNcAMax,
       P_NcAPosDiff := pNcAPosDiff,  P_NcAVeloDiff := pNcAVeloDiff,
       P_DrvSBip := pDrvSBip,  P_DrvSPos := pDrvSPos,
       P_DrvSNeg := pDrvSNeg,  P_DrvABip := pDrvABip,
       P_DrvAPos := pDrvAPos,  P_DrvANeg := pDrvANeg);
// done latches (Done is a single-scan pulse)
IF refPls.Done THEN dRef := TRUE; END_IF;
IF absDet.Done THEN dAbsD := TRUE; END_IF;
IF absSw.Done THEN dAbsS := TRUE; END_IF;
IF limSw.Done THEN dLim := TRUE; END_IF;
IF blk.Done THEN dBlk := TRUE; END_IF;
IF blkDet.Done THEN dBlkD := TRUE; END_IF;
IF blkLag.Done THEN dBlkL := TRUE; END_IF;
IF homeDir.Done THEN dHomeD := TRUE; END_IF;
IF finH.Done THEN dFin := TRUE; END_IF;
IF abortH.Done THEN dAbort := TRUE; END_IF;
IF flySw.Done THEN dFly := TRUE; END_IF;

// latch single-scan error outputs
IF refPls2.Error THEN errId1 := refPls2.ErrorID; END_IF;
IF refPls3.Error THEN errId2 := refPls3.ErrorID; END_IF;

// ---- stages ----------------------------------------------------------
IF st = 0 THEN
    ax.UNITS_PER_REV := 1000;
    ax.MAX_VEL := 100000;
    ax.MAX_ACCEL := 200000;
    ax.MAX_DECEL := 200000;
    ax.POS_MIN := -20000;
    ax.POS_MAX := 30000;
    ax.HOME_OFFSET := 0;
    ax.FOLLOW_WINDOW := 3;
    ax.FLAGS := 1;
    ax.OP := 1; ax();
    IF ax.AXIS <> 0 THEN axM := ax.AXIS; END_IF;
    IF axM <> 0 THEN
        mask := mask + 1;                          // bit0
        // pos-limit objects (sim ext): needed on the IO backend
        // where axis create does not carry the config struct
        ax.AXIS := axM;
        ax.OP := 5; ax.INDEX := 16#200A; ax.VALUE := -20000; ax();
        ax.OP := 5; ax.INDEX := 16#200B; ax.VALUE := 30000;  ax();
        ax.OP := 5; ax.INDEX := 16#200C; ax.VALUE := 1;      ax();
    END_IF;
    st := 1;
ELSIF st = 1 THEN
    IF pwr.Status THEN mask := mask + 2; st := 2; END_IF;
ELSIF st = 2 THEN
    IF sp.Done THEN mask := mask + 4; st := 3; END_IF;
ELSIF st = 3 THEN st := 4;
ELSIF st = 4 THEN st := 5;
ELSIF st = 5 THEN
    IF dRef AND ABS(posL - 100.0) < 5.0 AND pStored = TRUE THEN
        mask := mask + 8; st := 6;
    END_IF;
ELSIF st = 6 THEN
    IF sp.Done THEN st := 7; END_IF;
ELSIF st = 7 THEN st := 8;
ELSIF st = 8 THEN st := 9;
ELSIF st = 9 THEN
    IF dAbsD AND absDet.RecordedPosition <= -2700.0
       AND absDet.RecordedPosition >= -3300.0 THEN
        mask := mask + 16; st := 10;
    END_IF;
ELSIF st = 10 THEN
    IF sp.Done THEN st := 11; END_IF;
ELSIF st = 11 THEN st := 12;
ELSIF st = 12 THEN st := 13;
ELSIF st = 13 THEN
    IF dAbsS AND ABS(posL - 500.0) < 5.0 THEN
        mask := mask + 32; st := 14;
    END_IF;
ELSIF st = 14 THEN
    IF sp.Done THEN st := 15; END_IF;
ELSIF st = 15 THEN st := 16;
ELSIF st = 16 THEN st := 17;
ELSIF st = 17 THEN
    IF dLim AND ABS(posL - (-500.0)) < 5.0 THEN
        mask := mask + 64; st := 18;
    END_IF;
ELSIF st = 18 THEN
    IF sp.Done THEN st := 19; END_IF;
ELSIF st = 19 THEN st := 20;
ELSIF st = 20 THEN st := 21;
ELSIF st = 21 THEN
    IF dBlk AND ABS(posL - 25000.0) < 5.0 THEN
        mask := mask + 128; st := 22;
    END_IF;
ELSIF st = 22 THEN
    IF sp.Done THEN st := 23; END_IF;
ELSIF st = 23 THEN st := 24;
ELSIF st = 24 THEN st := 25;
ELSIF st = 25 THEN
    IF dBlkD AND blkDet.RecordedPosition <= -19000.0
       AND blkDet.RecordedPosition >= -21000.0 THEN
        mask := mask + 256; st := 26;
    END_IF;
ELSIF st = 26 THEN
    IF sp.Done THEN st := 27; END_IF;
ELSIF st = 27 THEN st := 28;
ELSIF st = 28 THEN st := 29;
ELSIF st = 29 THEN
    IF dBlkL AND ABS(posL - 20000.0) < 5.0 THEN
        mask := mask + 512; st := 30;
    END_IF;
ELSIF st = 30 THEN st := 31;
ELSIF st = 31 THEN
    IF dHomeD AND ABS(posL - 777.0) < 5.0 THEN
        mask := mask + 1024; st := 32;
    END_IF;
ELSIF st = 32 THEN st := 33;
ELSIF st = 33 THEN
    IF dFin AND ABS(posL - 1277.0) < 60.0
       AND pStored = FALSE THEN
        mask := mask + 2048; st := 34;
    END_IF;
ELSIF st = 34 THEN st := 35;
ELSIF st = 35 THEN
    IF dAbort THEN mask := mask + 4096; st := 36; END_IF;
ELSIF st = 36 THEN st := 37;
ELSIF st = 37 THEN st := 38;
ELSIF st = 38 THEN st := 39;
ELSIF st = 39 THEN
    IF dFly AND posL >= 4242.0 AND posL <= 4800.0 THEN
        mask := mask + 8192; st := 40;
    END_IF;
ELSIF st = 40 THEN st := 41;
ELSIF st = 41 THEN st := 42;
ELSIF st = 42 THEN st := 43;
ELSIF st = 43 THEN st := 44;
ELSIF st = 44 THEN
    IF errId1 = 16#4B93 THEN mask := mask + 16384; END_IF;
    st := 45;
ELSIF st = 45 THEN st := 46;
ELSIF st = 46 THEN
    IF errId2 = 16#4B91 THEN mask := mask + 32768; END_IF;
    st := 47;
END_IF;
END_PROGRAM

(* ---- tc3_mc3cam_case.st ---- *)
PROGRAM Tc3Mc3CamCase
VAR
    mask   AT %QD0 : DINT;
    st     : INT;
    prevSt : INT;
    pulse  : BOOL;
    started : BOOL;
    axM    : UDINT;
    axS    : UDINT;
    crM    : FB_MotionAxis;
    crS    : FB_MotionAxis;
    rdM    : FB_MotionAxis;
    wrM    : FB_MotionAxis;
    wrS    : FB_MotionAxis;
    pwrM   : MC_Power;
    pwrS   : MC_Power;
    phA    : MC_PhasingAbsolute;
    phR    : MC_PhasingRelative;
    gip    : MC_GearInPos;
    hph    : MC_HaltPhasing;
    mpos   : DINT;
    spos   : DINT;
    dPhA   : BOOL;
    dPhR   : BOOL;
    dGip   : BOOL;
    dHph   : BOOL;
    gipOff : BOOL;
    phEx   : BOOL;
    relEx  : BOOL;
    gipEx  : BOOL;
    hphEx  : BOOL;
END_VAR

pulse := FALSE;
IF NOT started THEN
    pulse := TRUE; started := TRUE;
ELSIF st <> prevSt THEN
    pulse := TRUE;
END_IF;
prevSt := st;

// per-scan position reads (diagnostic only; FBs do their own)
IF axM <> 0 THEN
    rdM.AXIS := axM; rdM.OP := 4; rdM.INDEX := 16#6064; rdM();
    mpos := rdM.VALUE;
END_IF;
IF axS <> 0 THEN
    rdM.AXIS := axS; rdM.OP := 4; rdM.INDEX := 16#6064; rdM();
    spos := rdM.VALUE;
END_IF;

// Execute is edge-triggered inside each FB; level-held here
phEx  := st = 2;
relEx := st = 4;
gipEx := st = 5;
hphEx := st = 6;

phA(Execute := phEx, PhaseShift := 5000, Velocity := 50000,
    Acceleration := 0, Deceleration := 0, Jerk := 0,
    Master := axM, Slave := axS);
phR(Execute := relEx, PhaseShift := 2000, Velocity := 50000,
    Acceleration := 0, Deceleration := 0, Jerk := 0,
    Master := axM, Slave := axS);
gip(Execute := gipEx, RatioNumerator := 1, RatioDenominator := 1,
    Velocity := 50000, Acceleration := 0, Deceleration := 0,
    Jerk := 0, Master := axM, Slave := axS);
hph(Execute := hphEx, Deceleration := 0, Jerk := 0,
    Master := axM, Slave := axS);

IF phA.Done THEN dPhA := TRUE; END_IF;
IF phR.Done THEN dPhR := TRUE; END_IF;
IF gip.InSync THEN dGip := TRUE; END_IF;
IF hph.Done THEN dHph := TRUE; END_IF;

IF st = 0 THEN
    crM.UNITS_PER_REV := 1000; crM.MAX_VEL := 100000;
    crM.MAX_ACCEL := 200000; crM.MAX_DECEL := 200000;
    crM.POS_MIN := -100000; crM.POS_MAX := 100000;
    crM.HOME_OFFSET := 0; crM.FOLLOW_WINDOW := 3; crM.FLAGS := 1;
    crM.OP := 1; crM();
    IF crM.AXIS <> 0 THEN axM := crM.AXIS; END_IF;
    crS.UNITS_PER_REV := 1000; crS.MAX_VEL := 100000;
    crS.MAX_ACCEL := 200000; crS.MAX_DECEL := 200000;
    crS.POS_MIN := -100000; crS.POS_MAX := 100000;
    crS.HOME_OFFSET := 0; crS.FOLLOW_WINDOW := 3; crS.FLAGS := 1;
    crS.OP := 1; crS();
    IF crS.AXIS <> 0 THEN axS := crS.AXIS; END_IF;
    IF axM <> 0 AND axS <> 0 THEN mask := mask + 1; END_IF; // bit0
    st := 1;
ELSIF st = 1 THEN
    pwrM(Enable := TRUE, Enable_Positive := TRUE,
         Enable_Negative := TRUE, Axis := axM);
    pwrS(Enable := TRUE, Enable_Positive := TRUE,
         Enable_Negative := TRUE, Axis := axS);
    IF pwrM.Status AND pwrS.Status THEN
        mask := mask + 2; st := 2;                     // bit1
    END_IF;
ELSIF st = 2 THEN
    // master: PV mode, constant velocity 20000 u/s; phA edge fires
    wrM.AXIS := axM; wrM.OP := 5; wrM.INDEX := 16#6060;
    wrM.VALUE := 3; wrM();
    wrM.OP := 5; wrM.INDEX := 16#60FF; wrM.VALUE := 20000; wrM();
    st := 3;
ELSIF st = 3 THEN
    // absolute phasing: slave must reach masterPos + 5000
    IF dPhA THEN
        mask := mask + 4; st := 4;                     // bit2
    END_IF;
ELSIF st = 4 THEN
    // relative phasing: +2000 additional phase on top of offset0
    IF dPhR THEN
        mask := mask + 8; st := 5;                     // bit3
    END_IF;
ELSIF st = 5 THEN
    // offset the slave +2000 once; gear-in-position must pull it
    // back onto the anchored trajectory
    IF NOT gipOff THEN
        gipOff := TRUE;
        wrS.AXIS := axS; wrS.OP := 5; wrS.INDEX := 16#6064;
        wrS.VALUE := spos + 2000; wrS();
    END_IF;
    IF dGip THEN
        mask := mask + 16; st := 6;                    // bit4
    END_IF;
ELSIF st = 6 THEN
    // halt phasing: slave ramps to rest
    IF dHph THEN
        mask := mask + 32; st := 7;                    // bit5
    END_IF;
ELSIF st = 7 THEN
    // hold; expect written at final step
END_IF;
END_PROGRAM

(* ---- tc3_mc3camtbl_case.st ---- *)
// tc3_mc3camtbl_case.st — Tc3_Mc3Camming cam-table e2e over the
// tplc-cam service: FB_CamTable object creation + WritePt/Config
// edges, MC_CamTableSelect, MC_CamIn CSP coupling (slave tracks
// master+5000 through an identity cam table), MC_CamScaling offset
// update, MC_ReadCamInfo and MC_CamRemove. Mask 0xff (8 checks).
PROGRAM Tc3Mc3CamTblCase
VAR
    mask   AT %QD0 : DINT;
    st     : INT;
    prevSt : INT;
    pulse  : BOOL;
    started : BOOL;
    wrN    : INT;
    axM    : UDINT;
    axS    : UDINT;
    camH   : UDINT;
    crM    : FB_MotionAxis;
    crS    : FB_MotionAxis;
    wrM    : FB_MotionAxis;
    wrS    : FB_MotionAxis;
    pwrM   : MC_Power;
    pwrS   : MC_Power;
    tbl    : FB_CamTable;
    camI   : MC_CamIn;
    camS   : MC_CamScaling;
    camSel : MC_CamTableSelect;
    camR   : MC_CamRemove;
    camInfo: MC_ReadCamInfo;
    dSel   : BOOL;
    dScl   : BOOL;
    dRem   : BOOL;
    dInfo1 : BOOL;
    dInfo2 : BOOL;
    iFound : UDINT;
    iCam   : UDINT;
    iMaster: UDINT;
    jFound : UDINT;
    gapSeen : BOOL;
    selEx  : BOOL;
    camInEx: BOOL;
    camScEx: BOOL;
    camRemEx: BOOL;
    infoEx : BOOL;
END_VAR

pulse := FALSE;
IF NOT started THEN
    pulse := TRUE; started := TRUE;
ELSIF st <> prevSt THEN
    pulse := TRUE;
END_IF;
prevSt := st;

// ---- level inputs, computed before the FB calls ----
tbl.WritePt := FALSE; tbl.ClearTable := FALSE; tbl.Config := FALSE;
IF st = 3 THEN
    IF wrN = 0 THEN
        tbl.PtIndex := 0; tbl.PtMaster := 0.0; tbl.PtSlave := 0.0;
        tbl.WritePt := TRUE;
    ELSIF wrN = 2 THEN
        tbl.PtIndex := 1; tbl.PtMaster := 100000.0;
        tbl.PtSlave := 100000.0; tbl.WritePt := TRUE;
    ELSIF wrN = 3 THEN
        tbl.Config := TRUE; tbl.TableCount := 2;
        tbl.Periodic := FALSE; tbl.Continuity := 0;
    END_IF;
END_IF

selEx := st = 5;
camInEx := st = 6;
camScEx := st = 7;
camRemEx := st = 9;
infoEx := (st = 7) OR (st = 9);

camI(Execute := camInEx, Master := axM, Slave := axS,
     CamObject := camH, SlaveOffset := 5000.0);
camS(Execute := camScEx, Slave := axS, CamObject := camH,
     SlaveOffset := 8000.0);
camSel(Execute := selEx, CamRef := camH, Periodic := FALSE,
       ContinuityRequirement := 0, CamObjectIn := camH);
camR(Execute := camRemEx, Slave := axS, CamObject := camH);
camInfo(Execute := infoEx, Slave := axS);
tbl();

IF camSel.Done THEN dSel := TRUE; END_IF;
IF camS.Done THEN dScl := TRUE; END_IF;
IF camR.Done THEN dRem := TRUE; END_IF;
IF camInfo.Done THEN
    IF st = 7 THEN
        dInfo1 := TRUE;
        iFound := camInfo.NumberOfCouplingsFound;
        iCam := camInfo.CamHandle;
        iMaster := camInfo.MasterAxis;
    ELSIF st = 9 THEN
        dInfo2 := TRUE;
        jFound := camInfo.NumberOfCouplingsFound;
    END_IF;
END_IF;

IF st = 0 THEN
    crM.UNITS_PER_REV := 1000; crM.MAX_VEL := 100000;
    crM.MAX_ACCEL := 200000; crM.MAX_DECEL := 200000;
    crM.POS_MIN := -100000; crM.POS_MAX := 100000;
    crM.HOME_OFFSET := 0; crM.FOLLOW_WINDOW := 3; crM.FLAGS := 1;
    crM.OP := 1; crM();
    IF crM.AXIS <> 0 THEN axM := crM.AXIS; END_IF;
    crS.UNITS_PER_REV := 1000; crS.MAX_VEL := 100000;
    crS.MAX_ACCEL := 200000; crS.MAX_DECEL := 200000;
    crS.POS_MIN := -100000; crS.POS_MAX := 100000;
    crS.HOME_OFFSET := 0; crS.FOLLOW_WINDOW := 3; crS.FLAGS := 1;
    crS.OP := 1; crS();
    IF crS.AXIS <> 0 THEN axS := crS.AXIS; END_IF;
    IF axM <> 0 AND axS <> 0 THEN mask := mask + 1; END_IF; // bit0
    st := 1;
ELSIF st = 1 THEN
    pwrM(Enable := TRUE, Enable_Positive := TRUE,
         Enable_Negative := TRUE, Axis := axM);
    pwrS(Enable := TRUE, Enable_Positive := TRUE,
         Enable_Negative := TRUE, Axis := axS);
    IF pwrM.Status AND pwrS.Status THEN
        mask := mask + 2; st := 2;                     // bit1
    END_IF;
ELSIF st = 2 THEN
    // master PV move; slave into CSP mode for 0x607A streaming
    wrM.AXIS := axM; wrM.OP := 5; wrM.INDEX := 16#6060;
    wrM.VALUE := 3; wrM();
    wrM.OP := 5; wrM.INDEX := 16#60FF; wrM.VALUE := 5000; wrM();
    wrS.AXIS := axS; wrS.OP := 5; wrS.INDEX := 16#6060;
    wrS.VALUE := 8; wrS();
    wrN := 0;
    st := 3;
ELSIF st = 3 THEN
    // cam table point writes + config (wrN sequencer, ~5 scans)
    wrN := wrN + 1;
    IF wrN >= 5 THEN st := 4; END_IF;
ELSIF st = 4 THEN
    IF tbl.Handle <> 0 THEN
        camH := tbl.Handle;
        mask := mask + 4; st := 5;                     // bit2
    END_IF;
ELSIF st = 5 THEN
    IF dSel THEN
        mask := mask + 8; st := 6;                     // bit3
    END_IF;
ELSIF st = 6 THEN
    // MC_CamIn bound on entry; slave must converge to mpos+5000
    IF camI.InSync THEN
        mask := mask + 16; st := 7;                    // bit4
    END_IF;
ELSIF st = 7 THEN
    // scaling update + cam info read
    IF dScl AND dInfo1 THEN
        IF iFound = 1 AND iCam = camH AND iMaster = axM THEN
            mask := mask + 32;                        // bit5
        END_IF;
        st := 8;
    END_IF;
ELSIF st = 8 THEN
    // wait for the +3000 target jump to break sync, then re-converge
    IF NOT camI.InSync THEN gapSeen := TRUE; END_IF;
    IF gapSeen AND camI.InSync THEN
        mask := mask + 64; st := 9;                    // bit6
    END_IF;
ELSIF st = 9 THEN
    // cam remove + second info read must show no coupling
    IF dRem AND dInfo2 THEN
        IF jFound = 0 THEN
            mask := mask + 128;                       // bit7
        END_IF;
        st := 10;
    END_IF;
ELSIF st = 10 THEN
    // hold; expect written at final step
END_IF;
END_PROGRAM

(* ---- tc3_mc3ptp_case.st ---- *)
PROGRAM Tc3Mc3PtpCase
VAR
    mask   AT %QD0 : DINT;
    st     : INT;
    prevSt : INT;
    pulse  : BOOL;
    started : BOOL;
    axM    : UDINT;
    ax     : FB_MotionAxis;
    rd     : FB_MotionAxis;
    pwr    : MC_Power;
    rst    : MC_Reset;
    tq     : MC_ReadActualTorque;
    hwr    : MC_WriteHardwareParameter;
    hrr    : MC_ReadHardwareParameter;
    wfs    : MC_WaitForStableActualPosition;
    te     : MC_TriggerError;
    hs     : MC_SetHomingState;
    lc     : MC_LoadControl;
    esg    : MC_ActivateExternalSetpointGeneration;
    axErr  : MC_ReadAxisError;
    vel    : DINT;
END_VAR

// per-scan snapshot
IF axM <> 0 THEN
    rd.AXIS := axM; rd.OP := 6; rd();
    vel := rd.VEL_ACTUAL;
END_IF;

pulse := FALSE;
IF NOT started THEN
    pulse := TRUE; started := TRUE;
ELSIF st <> prevSt THEN
    pulse := TRUE;
END_IF;
prevSt := st;

IF st = 0 THEN
    ax.UNITS_PER_REV := 1000;
    ax.MAX_VEL := 100000;
    ax.MAX_ACCEL := 200000;
    ax.MAX_DECEL := 200000;
    ax.POS_MIN := -20000;
    ax.POS_MAX := 30000;
    ax.HOME_OFFSET := 0;
    ax.FOLLOW_WINDOW := 3;
    ax.FLAGS := 1;
    ax.OP := 1; ax();
    IF ax.AXIS <> 0 THEN axM := ax.AXIS; END_IF;
    IF axM <> 0 THEN mask := mask + 1; END_IF;   // bit0: create
    st := 1;
ELSIF st = 1 THEN
    pwr(Enable := TRUE, Enable_Positive := TRUE,
        Enable_Negative := TRUE, Axis := axM);
    IF pwr.Status THEN mask := mask + 2; st := 2; END_IF;  // bit1: power
ELSIF st = 2 THEN
    tq(Enable := TRUE, Axis := axM);
    hwr(Execute := pulse, ParameterNumber := 16#6065,
        Value := 5, Axis := axM);
    IF pulse AND hwr.Done AND tq.Valid THEN
        mask := mask + 4;                        // bit2: torque+hw wr
    END_IF;
    st := 3;
ELSIF st = 3 THEN
    hrr(Enable := TRUE, ParameterNumber := 16#6065, Axis := axM);
    IF hrr.Valid AND hrr.Value = 5 THEN
        mask := mask + 8;                        // bit3: hw param rd
    END_IF;
    st := 4;
ELSIF st = 4 THEN
    wfs(Execute := pulse, PositionWindow := 10,
        VelocityWindow := 1, Axis := axM);
    IF wfs.Done THEN mask := mask + 16; st := 5; END_IF;  // bit4: stable
ELSIF st = 5 THEN
    hs(Execute := pulse, HomingState := 1, Axis := axM);
    lc(Execute := pulse, Axis := axM);
    esg(Execute := pulse, Axis := axM);
    IF pulse AND hs.Done AND lc.Done AND esg.Done THEN
        mask := mask + 32;                       // bit5: no-op FBs
    END_IF;
    st := 6;
ELSIF st = 6 THEN
    te(Execute := pulse, ErrorCode := 4660, Axis := axM); // 0x1234
    IF pulse AND te.Done THEN mask := mask + 64; st := 7; END_IF; // bit6
ELSIF st = 7 THEN
    axErr(Enable := TRUE, Axis := axM);
    IF axErr.Valid AND axErr.AxisErrorID = 4660 THEN
        mask := mask + 128;                      // bit7: fault latched
    END_IF;
    rst(Execute := pulse, Axis := axM);
    IF pulse AND rst.Done THEN st := 8; END_IF;
ELSIF st = 8 THEN
    axErr(Enable := TRUE, Axis := axM);
    IF axErr.Valid AND axErr.AxisErrorID = 0 THEN
        mask := mask + 256;                      // bit8: fault cleared
    END_IF;
    st := 9;
ELSIF st = 9 THEN
    // hold; expect written at final step
END_IF;
END_PROGRAM

(* ---- tc3_mcgroup_case.st ---- *)
PROGRAM Tc3McGroupCase
VAR
    mask   AT %QD0 : DINT;
    st     : INT;
    prevSt : INT;
    cur    : INT;
    pulse  : BOOL;
    started : BOOL;
    grp    : UDINT;
    grpBad : UDINT;
    ax7    : UDINT;
    ax9    : UDINT;
    addA   : MC_AddAxisToGroup;
    addB   : MC_AddAxisToGroup;
    remA   : MC_RemoveAxisFromGroup;
    ungrp  : MC_UngroupAllAxes;
    enA    : MC_GroupEnable;
    enBad  : MC_GroupEnable;
    disA   : MC_GroupDisable;
    rstA   : MC_GroupReset;
    rs     : MC_GroupReadStatus;
    re     : MC_GroupReadError;
    so     : MC_GroupSetOverride;
    ss     : MC_GroupSetSetpointSource;
    ct     : MC_SetCoordinateTransform;
    ident  : UDINT;
    mg     : FB_McGroup;
    memOk  : BOOL;
END_VAR

cur := st;
pulse := (cur <> prevSt) OR NOT started;
started := TRUE;
prevSt := cur;

grp := 1;
grpBad := 2;
ax7 := 7;
ax9 := 9;
ident := UDINT_TO_IDENTINGROUP(0);
memOk := FALSE;

// Level-triggered readers: called every scan.
rs(Enable := TRUE, AxesGroup := grp);
re(Enable := TRUE, AxesGroup := grp);

// st0: add axis 7 to group 1 (ident 0)
IF cur = 0 THEN
    addA(Execute := pulse, IdentInGroup := ident,
         AxesGroup := grp, Axis := ax7);
    IF pulse AND addA.Done AND NOT addA.Error THEN
        mask := mask + 1;                       // bit0: add axis
    END_IF;
    st := 1;
// st1: status readback -> disabled, valid
ELSIF cur = 1 THEN
    IF rs.Valid AND rs.GroupDisabled THEN
        mask := mask + 2;                       // bit1: read status
    END_IF;
    st := 2;
// st2: enable group -> standby
ELSIF cur = 2 THEN
    enA(Execute := pulse, AxesGroup := grp);
    IF pulse AND enA.Done AND NOT enA.Error THEN
        mask := mask + 4;                       // bit2: enable done
    END_IF;
    st := 3;
// st3: status now standby + group error read valid
ELSIF cur = 3 THEN
    IF rs.GroupStandby AND re.Valid AND re.GroupErrorId = 0 THEN
        mask := mask + 8;                       // bit3: standby+err
    END_IF;
    st := 4;
// st4: enable empty group 2 -> error
ELSIF cur = 4 THEN
    enBad(Execute := pulse, AxesGroup := grpBad);
    IF pulse AND enBad.Error THEN
        mask := mask + 16;                      // bit4: empty enable err
    END_IF;
    st := 5;
// st5: override 150%
ELSIF cur = 5 THEN
    so(Execute := pulse, Enable := TRUE, VelFactor := 1.5,
       AxesGroup := grp);
    IF pulse AND so.Done AND
       ABS(so.OverrideActual - 1.5) < 0.001 THEN
        mask := mask + 32;                      // bit5: override
    END_IF;
    st := 6;
// st6: setpoint source MCS (2)
ELSIF cur = 6 THEN
    ss(Execute := pulse, SetpointSource := 2, AxesGroup := grp);
    IF pulse AND ss.Done AND NOT ss.Error THEN
        mask := mask + 64;                      // bit6: setpoint src
    END_IF;
    st := 7;
// st7: coordinate transform 3 -> active
ELSIF cur = 7 THEN
    ct(Execute := pulse, CoordTransform := 3, AxesGroup := grp);
    IF pulse AND ct.Done AND ct.Active AND NOT ct.Error THEN
        mask := mask + 128;                     // bit7: coord transform
    END_IF;
    st := 8;
// st8: membership readback via raw FB_McGroup OP10
ELSIF cur = 8 THEN
    mg.OP := 10; mg.GRP := grp; mg();
    IF mg.STATUS = 0 AND mg.NAXES = 1 AND mg.AXES[0] = 7 THEN
        memOk := TRUE;
        mask := mask + 256;                     // bit8: membership
    END_IF;
    st := 9;
// st9: disable group (membership changes need disabled state)
ELSIF cur = 9 THEN
    disA(Execute := pulse, AxesGroup := grp);
    IF pulse AND disA.Done THEN st := 10; END_IF;
// st10: add axis 9, remove axis 7 -> still 1 member (9)
ELSIF cur = 10 THEN
    addB(Execute := pulse, IdentInGroup := ident,
         AxesGroup := grp, Axis := ax9);
    remA(Execute := pulse, IdentInGroup := ident,
          AxesGroup := grp, Axis := ax7);
    IF pulse AND addB.Done AND remA.Done THEN st := 11; END_IF;
// st11: verify swap + ungroup all
ELSIF cur = 11 THEN
    mg.OP := 10; mg.GRP := grp; mg();
    IF mg.STATUS = 0 AND mg.NAXES = 1 AND mg.AXES[0] = 9 THEN
        mask := mask + 512;                     // bit9: swap member
    END_IF;
    ungrp(Execute := pulse, AxesGroup := grp);
    IF pulse AND ungrp.Done AND NOT ungrp.Error THEN
        mask := mask + 1024;                    // bit10: ungroup
    END_IF;
    st := 12;
// st12: group reset on fresh group
ELSIF cur = 12 THEN
    rstA(Execute := pulse, AxesGroup := grpBad);
    IF pulse AND rstA.Done THEN
        mask := mask + 2048;                    // bit11: reset
    END_IF;
    st := 13;
ELSIF cur = 13 THEN
    // hold; expect written at final step
END_IF;
END_PROGRAM

(* ---- tc3_mcgroup_stop_case.st ---- *)
// tc3_mcgroup_stop_case.st — Tc3_McCoordinatedMotion group motion
// e2e: two real axes grouped via MC_AddAxisToGroup, PV velocity
// moves, then MC_GroupStop (ramp to rest) and MC_GroupHalt
// (immediate disable) with per-axis VEL_ACTUAL verification.
// Mask 0x3f (6 checks).
PROGRAM Tc3McGroupStopCase
VAR
    mask   AT %QD0 : DINT;
    st     : INT;
    prevSt : INT;
    pulse  : BOOL;
    started : BOOL;
    dwell  : INT;
    grp    : UDINT := 1;
    axA    : UDINT;
    axB    : UDINT;
    crA    : FB_MotionAxis;
    crB    : FB_MotionAxis;
    rdA    : FB_MotionAxis;
    rdB    : FB_MotionAxis;
    wrA    : FB_MotionAxis;
    wrB    : FB_MotionAxis;
    pwrA   : MC_Power;
    pwrB   : MC_Power;
    addA   : MC_AddAxisToGroup;
    addB   : MC_AddAxisToGroup;
    gStop  : MC_GroupStop;
    gHalt  : MC_GroupHalt;
    vA     : DINT;
    vB     : DINT;
    dAddA  : BOOL;
    dAddB  : BOOL;
    dStop  : BOOL;
    dHalt  : BOOL;
    gStopEx: BOOL;
    gHaltEx: BOOL;
END_VAR

pulse := FALSE;
IF NOT started THEN
    pulse := TRUE; started := TRUE;
ELSIF st <> prevSt THEN
    pulse := TRUE; dwell := 0;
END_IF;
prevSt := st;

// per-scan velocity reads
IF axA <> 0 THEN
    rdA.AXIS := axA; rdA.OP := 3; rdA();
    rdA.OP := 4; rdA.INDEX := 16#606C; rdA(); vA := rdA.VALUE;
END_IF;
IF axB <> 0 THEN
    rdB.AXIS := axB; rdB.OP := 3; rdB();
    rdB.OP := 4; rdB.INDEX := 16#606C; rdB(); vB := rdB.VALUE;
END_IF;

gStopEx := st = 6;
gHaltEx := st = 10;
gStop(Execute := gStopEx, Deceleration := 1000.0, AxesGroup := grp);
gHalt(Execute := gHaltEx, AxesGroup := grp);

IF gStop.Done THEN dStop := TRUE; END_IF;
IF gHalt.Done THEN dHalt := TRUE; END_IF;

IF st = 0 THEN
    crA.UNITS_PER_REV := 1000; crA.MAX_VEL := 100000;
    crA.MAX_ACCEL := 200000; crA.MAX_DECEL := 200000;
    crA.POS_MIN := -100000; crA.POS_MAX := 100000;
    crA.HOME_OFFSET := 0; crA.FOLLOW_WINDOW := 3; crA.FLAGS := 1;
    crA.OP := 1; crA();
    IF crA.AXIS <> 0 THEN axA := crA.AXIS; END_IF;
    crB.UNITS_PER_REV := 1000; crB.MAX_VEL := 100000;
    crB.MAX_ACCEL := 200000; crB.MAX_DECEL := 200000;
    crB.POS_MIN := -100000; crB.POS_MAX := 100000;
    crB.HOME_OFFSET := 0; crB.FOLLOW_WINDOW := 3; crB.FLAGS := 1;
    crB.OP := 1; crB();
    IF crB.AXIS <> 0 THEN axB := crB.AXIS; END_IF;
    IF axA <> 0 AND axB <> 0 THEN mask := mask + 1; END_IF; // bit0
    st := 1;
ELSIF st = 1 THEN
    pwrA(Enable := TRUE, Enable_Positive := TRUE,
         Enable_Negative := TRUE, Axis := axA);
    pwrB(Enable := TRUE, Enable_Positive := TRUE,
         Enable_Negative := TRUE, Axis := axB);
    IF pwrA.Status AND pwrB.Status THEN
        mask := mask + 2; st := 2;                     // bit1
    END_IF;
ELSIF st = 2 THEN
    // add axis A to a fresh group (ensure creates the handle)
    addA(Execute := pulse, IdentInGroup := 0,
         AxesGroup := grp, Axis := axA);
    IF addA.Done THEN dAddA := TRUE; END_IF;
    IF dAddA THEN st := 3; END_IF;
ELSIF st = 3 THEN
    addB(Execute := pulse, IdentInGroup := 0,
         AxesGroup := grp, Axis := axB);
    IF addB.Done THEN dAddB := TRUE; END_IF;
    IF dAddB THEN
        mask := mask + 4; st := 4;                     // bit2
    END_IF;
ELSIF st = 4 THEN
    // both axes: PV mode, velocity 5000 u/s
    wrA.AXIS := axA; wrA.OP := 5; wrA.INDEX := 16#6060;
    wrA.VALUE := 3; wrA();
    wrA.OP := 5; wrA.INDEX := 16#60FF; wrA.VALUE := 5000; wrA();
    wrB.AXIS := axB; wrB.OP := 5; wrB.INDEX := 16#6060;
    wrB.VALUE := 3; wrB();
    wrB.OP := 5; wrB.INDEX := 16#60FF; wrB.VALUE := 5000; wrB();
    st := 5;
ELSIF st = 5 THEN
    // let both axes spin up, then confirm motion
    dwell := dwell + 1;
    IF dwell >= 15 THEN
        IF vA > 0 AND vB > 0 THEN
            mask := mask + 8;                         // bit3
        END_IF;
        st := 6;
    END_IF;
ELSIF st = 6 THEN
    // group stop: ramp to rest; Done implies all VEL_ACTUAL = 0
    IF dStop THEN
        mask := mask + 16; st := 7;                    // bit4
    END_IF;
ELSIF st = 7 THEN
    // restart both axes for the halt test
    wrA.AXIS := axA; wrA.OP := 5; wrA.INDEX := 16#6060;
    wrA.VALUE := 3; wrA();
    wrA.OP := 5; wrA.INDEX := 16#60FF; wrA.VALUE := 5000; wrA();
    wrB.AXIS := axB; wrB.OP := 5; wrB.INDEX := 16#6060;
    wrB.VALUE := 3; wrB();
    wrB.OP := 5; wrB.INDEX := 16#60FF; wrB.VALUE := 5000; wrB();
    st := 8;
ELSIF st = 8 THEN
    dwell := dwell + 1;
    IF dwell >= 15 THEN st := 10; END_IF;
ELSIF st = 10 THEN
    // group halt: immediate disable; Done implies all stopped
    IF dHalt THEN
        mask := mask + 32; st := 11;                   // bit5
    END_IF;
ELSIF st = 11 THEN
    // hold; expect written at final step
END_IF;
END_PROGRAM

(* ---- tc3_mcpath_case.st ---- *)
// tc3_mcpath_case.st — Tc3_McCoordinatedMotion path e2e: two real
// axes grouped, a 3-segment path (linear -> dwell -> linear)
// prepared through MC_MoveLinearAbsolutePreparation /
// MC_DwellTimePreparation, executed by MC_MovePath with per-scan
// 0x607A CSP streaming, final-position verification.
// Mask 0x3f (6 checks).
PROGRAM Tc3McPathCase
VAR
    mask   AT %QD0 : DINT;
    st     : INT;
    prevSt : INT;
    pulse  : BOOL;
    started : BOOL;
    grp    : UDINT := 1;
    pathH  : UDINT := 0;
    axA    : UDINT;
    axB    : UDINT;
    crA    : FB_MotionAxis;
    crB    : FB_MotionAxis;
    rdA    : FB_MotionAxis;
    rdB    : FB_MotionAxis;
    pwrA   : MC_Power;
    pwrB   : MC_Power;
    addA   : MC_AddAxisToGroup;
    addB   : MC_AddAxisToGroup;
    prep1  : MC_MoveLinearAbsolutePreparation;
    prepD  : MC_DwellTimePreparation;
    prepB  : MC_MoveBlendingPreparation;
    prepK  : MC_BlockerPreparation;
    relBlk : MC_ReleaseBlocker;
    blkSt  : MC_GroupReadBlockerStatus;
    trajRd : MC_GroupReadTrajectoryInformation;
    trafoPrep : MC_SetCoordinateTransformPreparation;
    setTrafo : MC_SetCoordinateTransform;
    mgRd   : FB_McGroup;
    prepC  : MC_MoveCircularAbsolutePreparation;
    prep2  : MC_MoveDirectPreparation;
    mvPath : MC_MovePath;
    pos1   : ARRAY[0..15] OF LREAL;
    pos2   : ARRAY[0..15] OF LREAL;
    auxC   : ARRAY[0..15] OF LREAL;
    endC   : ARRAY[0..15] OF LREAL;
    transP : ARRAY[0..15] OF LREAL;
    dAddA  : BOOL;
    dAddB  : BOOL;
    dPrep1 : BOOL;
    dPrepD : BOOL;
    dPrep2 : BOOL;
    dPath  : BOOL;
    busySeen : BOOL;
    gotBusy : BOOL;
    gotPos  : BOOL;
    sawBlocked : BOOL;
    sawTraj : BOOL;
    coordNow : UDINT;
    mCnt   : INT;
    dRel   : BOOL;
    pA     : DINT;
    pB     : DINT;
END_VAR

pulse := FALSE;
IF NOT started THEN
    pulse := TRUE; started := TRUE;
ELSIF st <> prevSt THEN
    pulse := TRUE;
END_IF;
prevSt := st;

// per-scan position reads
IF axA <> 0 THEN
    rdA.AXIS := axA; rdA.OP := 4; rdA.INDEX := 16#6064; rdA(); pA := rdA.VALUE;
END_IF;
IF axB <> 0 THEN
    rdB.AXIS := axB; rdB.OP := 4; rdB.INDEX := 16#6064; rdB(); pB := rdB.VALUE;
END_IF;

mvPath(Execute := st = 8, AxesGroup := grp, PathData := pathH);
IF mvPath.Busy THEN busySeen := TRUE; END_IF;
IF mvPath.Done THEN dPath := TRUE; END_IF;

IF st = 0 THEN
    crA.UNITS_PER_REV := 1000; crA.MAX_VEL := 100000;
    crA.MAX_ACCEL := 200000; crA.MAX_DECEL := 200000;
    crA.POS_MIN := -100000; crA.POS_MAX := 100000;
    crA.HOME_OFFSET := 0; crA.FOLLOW_WINDOW := 3; crA.FLAGS := 1;
    crA.OP := 1; crA();
    IF crA.AXIS <> 0 THEN axA := crA.AXIS; END_IF;
    crB.UNITS_PER_REV := 1000; crB.MAX_VEL := 100000;
    crB.MAX_ACCEL := 200000; crB.MAX_DECEL := 200000;
    crB.POS_MIN := -100000; crB.POS_MAX := 100000;
    crB.HOME_OFFSET := 0; crB.FOLLOW_WINDOW := 3; crB.FLAGS := 1;
    crB.OP := 1; crB();
    IF crB.AXIS <> 0 THEN axB := crB.AXIS; END_IF;
    IF axA <> 0 AND axB <> 0 THEN mask := mask + 1; END_IF; // bit0
    st := 1;
ELSIF st = 1 THEN
    pwrA(Enable := TRUE, Enable_Positive := TRUE,
         Enable_Negative := TRUE, Axis := axA);
    pwrB(Enable := TRUE, Enable_Positive := TRUE,
         Enable_Negative := TRUE, Axis := axB);
    IF pwrA.Status AND pwrB.Status THEN
        mask := mask + 2; st := 2;                     // bit1
    END_IF;
ELSIF st = 2 THEN
    addA(Execute := pulse, IdentInGroup := 0,
         AxesGroup := grp, Axis := axA);
    IF addA.Done THEN dAddA := TRUE; END_IF;
    IF dAddA THEN st := 3; END_IF;
ELSIF st = 3 THEN
    addB(Execute := pulse, IdentInGroup := 0,
         AxesGroup := grp, Axis := axB);
    setTrafo(Execute := pulse, CoordTransform := 3,
             AxesGroup := grp);
    IF addB.Done THEN dAddB := TRUE; END_IF;
    IF dAddB THEN
        mask := mask + 4; st := 4;                     // bit2
    END_IF;
ELSIF st = 4 THEN
    // segment 1: linear to (1000, 0)
    pos1[0] := 1000.0; pos1[1] := 0.0;
    prep1(Execute := pulse, Position := pos1, PositionCount := 2,
          Velocity := 20000.0, Acceleration := 50000.0,
          Deceleration := 50000.0, Jerk := 0.0, BufferMode := 1,
          PathData := pathH);
    IF prep1.Error THEN mask := mask + 256; END_IF;
    IF NOT prep1.Error THEN dPrep1 := TRUE; END_IF;
    IF dPrep1 THEN st := 5; END_IF;
ELSIF st = 5 THEN
    // segment 2: circular, center (0,0), end (0,1000), CCW
    auxC[0] := 0.0; auxC[1] := 0.0;
    endC[0] := 0.0; endC[1] := 1000.0;
    prepC(Execute := pulse, CircMode := 1,
          AuxPoint := auxC, AuxPointCount := 2,
          EndPoint := endC, EndPointCount := 2,
          PathChoice := 1, Velocity := 20000.0,
          Acceleration := 50000.0, Deceleration := 50000.0,
          Jerk := 0.0, BufferMode := 1, PathData := pathH);
    IF prepC.Error THEN mask := mask + 256; END_IF;
    IF NOT prepC.Error THEN dPrepD := TRUE; END_IF;
    IF dPrepD THEN st := 6; END_IF;
ELSIF st = 6 THEN
    // segment 3: dwell 200 ms, then a 150 ms blend junction
    prepD(Execute := pulse, DwellTime := 200, BufferMode := 1,
          PathData := pathH);
    transP[0] := 150.0;
    prepB(Execute := pulse, Velocity := 20000.0,
          Acceleration := 50000.0, Deceleration := 50000.0,
          Jerk := 0.0, BufferMode := 1, TransitionMode := 0,
          TransitionParameter := transP,
          TransitionParameterCount := 1, InvokeId := 0,
          PathData := pathH);
    IF prepD.Error OR prepB.Error THEN mask := mask + 256; END_IF;
    IF NOT prepD.Error AND NOT prepB.Error THEN st := 7; END_IF;
ELSIF st = 7 THEN
    // transform marker -> coord 9, blocker gate id 7, linear
    trafoPrep(PathData := pathH, CoordTransform := 9);
    prepK(Execute := pulse, BlockerId := 7, BufferMode := 1,
          PathData := pathH);
    pos2[0] := 2000.0; pos2[1] := 2000.0;
    prep2(Execute := pulse, Position := pos2, PositionCount := 2,
          Velocity := 20000.0, Acceleration := 50000.0,
          Deceleration := 50000.0, Jerk := 0.0, BufferMode := 1,
          PathData := pathH);
    IF prepK.Error OR prep2.Error THEN mask := mask + 256; END_IF;
    IF NOT prepK.Error AND NOT prep2.Error THEN dPrep2 := TRUE; END_IF;
    IF dPrep2 THEN
        // 6 segments prepared on a live path handle
        IF pathH <> 0 THEN mask := mask + 8; END_IF;   // bit3
        st := 8;
    END_IF;
ELSIF st = 8 THEN
    // path running; blocker status polled, release after ~1.2 s
    blkSt(Enable := TRUE, AxesGroup := grp);
    IF blkSt.Blocked THEN sawBlocked := TRUE; END_IF;
    trajRd(Enable := TRUE, AxesGroup := grp);
    IF trajRd.Valid AND trajRd.EntryCount >= 3 THEN
        sawTraj := TRUE;
    END_IF;
    IF busySeen THEN gotBusy := TRUE; END_IF;
    mCnt := mCnt + 1;
    IF mCnt >= 120 THEN st := 9; END_IF;
ELSIF st = 9 THEN
    // release the blocker gate
    relBlk(Execute := pulse, BlockerId := 7, AxesGroup := grp);
    IF relBlk.Done THEN dRel := TRUE; END_IF;
    IF dRel THEN st := 10; END_IF;
ELSIF st = 10 THEN
    // path resumes and finishes
    IF dPath THEN
        // final positions near (2000, 2000), tolerance 300, and the
        // coordinate transform must have switched to 9 mid-path
        mgRd.GRP := grp; mgRd.OP := 11; mgRd();
        coordNow := mgRd.COORD;
        IF ABS(pA - 2000) < 300 AND ABS(pB - 2000) < 300 AND
           coordNow = 9 THEN
            gotPos := TRUE;
        END_IF;
        IF gotBusy THEN mask := mask + 16; END_IF;   // bit4
        IF gotPos THEN mask := mask + 32; END_IF;    // bit5
        IF sawBlocked THEN mask := mask + 64; END_IF; // bit6
        IF sawTraj THEN mask := mask + 128; END_IF;  // bit7
        st := 11;
    END_IF;
ELSIF st = 11 THEN
    // hold; expect written at final step
END_IF;
END_PROGRAM
